REGION Network 14: 关门停止控制
   // 1.脚踢开关又有信号
   // 2.操作门关位有信号
   // 3.操作门关门时间超时
   // 4.门电机保护有信号
   // 5.再次点击开门触摸按钮
   // 6.再次点击关门触摸按钮
   // 7.再次点击机械开门按钮
   // 8.再次点击机械关门按钮
   // 9..操作门有障碍
   RUNG wire#powerrail
      { S7_Templates := "SrcType := Word" } EQ_Contact(in1 := #门状态, in2 := 2)
      wire#w1
      Contact( #脚踢开关状态 )
      wire#w2
      Move(in := 0, out1 => #门状态)
      wire#w3
      R_Coil( #触摸开门按钮状态 )
      R_Coil( #机械开门按钮状态 )
      R_Coil( #机械关门按钮状态 )
      R_Coil( #脚踢开关状态 )
      R_Coil( #触摸关门按钮状态 )
   END_RUNG
   RUNG wire#w1
      Contact( #操作门关位 )
   END_RUNG wire#w2
   RUNG wire#w1
      { S7_Templates := "SrcType := UInt" } GT_Contact(in1 := #关门时间统计, in2 := #操作门最大关闭时间秒)
   END_RUNG wire#w2
   RUNG wire#w1
      Contact( #门电机保护信号 )
   END_RUNG wire#w2
   RUNG wire#w1
      Contact( #机械开门按钮状态 )
   END_RUNG wire#w2
   RUNG wire#w1
      Contact( #机械关门按钮状态 )
   END_RUNG wire#w2
   RUNG wire#w1
      Contact( #触摸关门按钮状态 )
   END_RUNG wire#w2
   RUNG wire#w1
      Contact( #触摸开门按钮状态 )
   END_RUNG wire#w2
   RUNG wire#w1
      I_Contact( #操作门障碍 )
   END_RUNG wire#w2
   RUNG wire#w3
      { S7_Templates := "SrcType := UInt" } GT_Contact(in1 := #关门时间统计, in2 := #操作门最大关闭时间秒)
      I_Contact( #报警开关.%X3 )
      S_Coil( #报警码.%X3 )
   END_RUNG
   RUNG wire#w3
      I_Contact( #操作门障碍 )
      wire#w4
      S_Coil( #关闭门失败后需要开门标志 )
      Move(in := 0, out1 => #门关闭失败重新开门等待时间)
   END_RUNG
   RUNG wire#w4
      I_Contact( #报警开关.%X5 )
      S_Coil( #报警码.%X5 )
   END_RUNG
   RUNG wire#w3
      Contact( #门电机保护信号 )
      I_Contact( #报警开关.%X4 )
      S_Coil( #报警码.%X4 )
   END_RUNG
   // the same network as SCL:
   #_w1 := (#门状态 = 2) AND (#脚踢开关状态 OR #操作门关位 OR (#关门时间统计 > #操作门最大关闭时间秒) OR #门电机保护信号 OR #机械开门按钮状态 OR #机械关门按钮状态 OR #触摸关门按钮状态 OR #触摸开门按钮状态 OR NOT #操作门障碍);
   IF #_w1 THEN
       #门状态 := 0;
       #触摸开门按钮状态 := FALSE;
       #机械开门按钮状态 := FALSE;
       #机械关门按钮状态 := FALSE;
       #脚踢开关状态 := FALSE;
       #触摸关门按钮状态 := FALSE;
   END_IF;
   IF #_w1 AND (#关门时间统计 > #操作门最大关闭时间秒) AND NOT #报警开关.%X3 THEN #报警码.%X3 := TRUE; END_IF;
   #_w2 := #_w1 AND NOT #操作门障碍;
   IF #_w2 THEN
       #关闭门失败后需要开门标志 := TRUE;
       #门关闭失败重新开门等待时间 := 0;
   END_IF;
   IF #_w2 AND NOT #报警开关.%X5 THEN #报警码.%X5 := TRUE; END_IF;
   IF #_w1 AND #门电机保护信号 AND NOT #报警开关.%X4 THEN #报警码.%X4 := TRUE; END_IF;
END_REGION

REGION Network 15: 如果是前门遇到障碍,门停止后,还需要将门打开
   // 关门失败后,门先停止0.8秒 然后再开门
   RUNG wire#powerrail
      { S7_Templates := "SrcType := Word" } EQ_Contact(in1 := #门状态, in2 := 0)
      Contact( #关闭门失败后需要开门标志 )
      wire#w1
      Contact( "Clock_10Hz" )
      P_Trig( #门关闭失败重新开门时间统计沿 )
      { S7_Templates := "DestType := UInt" } Inc( #门关闭失败重新开门等待时间 )
   END_RUNG
   RUNG wire#w1
      { S7_Templates := "SrcType := UInt" } GE_Contact(in1 := #门关闭失败重新开门等待时间, in2 := 8)
      wire#w2
      S_Coil( #触摸开门按钮状态 )
   END_RUNG
   RUNG wire#w2
      R_Coil( #关闭门失败后需要开门标志 )
      Move(in := 0, out1 => #门关闭失败重新开门等待时间)
   END_RUNG
   // the same network as SCL:
   #_w1 := (#门状态 = 0) AND #关闭门失败后需要开门标志;
   #_w2 := #_w1 AND "Clock_10Hz";
   #_w3 := #_w2 AND NOT #门关闭失败重新开门时间统计沿;   // rising edge
   #门关闭失败重新开门时间统计沿 := #_w2;
   IF #_w3 THEN #门关闭失败重新开门等待时间 := #门关闭失败重新开门等待时间 + 1; END_IF;
   IF #_w1 AND (#门关闭失败重新开门等待时间 >= 8) THEN
       #触摸开门按钮状态 := TRUE;
       #关闭门失败后需要开门标志 := FALSE;
       #门关闭失败重新开门等待时间 := 0;
   END_IF;
END_REGION

REGION Network 16: 其他门报警
   // 1.同时检测到操作门关位和开位1秒
   RUNG wire#powerrail
      Contact( #操作门开位 )
      Contact( #操作门关位 )
      wire#w1
      Contact( "Clock_10Hz" )
      P_Trig( #同时检测到门开关位时间统计沿 )
      { S7_Templates := "DestType := UInt" } Inc( #同时检测到门开位和关位信号时间统计 )
   END_RUNG
   RUNG wire#w1
      { S7_Templates := "SrcType := UInt" } GE_Contact(in1 := #同时检测到门开位和关位信号时间统计, in2 := 10)
      Move(in := 10, out1 => #同时检测到门开位和关位信号时间统计)
      I_Contact( #报警开关.%X6 )
      S_Coil( #报警码.%X6 )
   END_RUNG
   RUNG wire#powerrail
      I_Contact( #操作门开位 )
      wire#w2
      Move(in := 0, out1 => #同时检测到门开位和关位信号时间统计)
   END_RUNG
   RUNG wire#powerrail
      I_Contact( #操作门关位 )
   END_RUNG wire#w2
   // the same network as SCL:
   #_w1 := #操作门开位 AND #操作门关位;
   #_w2 := #_w1 AND "Clock_10Hz";
   #_w3 := #_w2 AND NOT #同时检测到门开关位时间统计沿;   // rising edge
   #同时检测到门开关位时间统计沿 := #_w2;
   IF #_w3 THEN #同时检测到门开位和关位信号时间统计 := #同时检测到门开位和关位信号时间统计 + 1; END_IF;
   #_w4 := #_w1 AND (#同时检测到门开位和关位信号时间统计 >= 10);
   IF #_w4 THEN #同时检测到门开位和关位信号时间统计 := 10; END_IF;
   IF #_w4 AND NOT #报警开关.%X6 THEN #报警码.%X6 := TRUE; END_IF;
   IF NOT #操作门开位 OR NOT #操作门关位 THEN #同时检测到门开位和关位信号时间统计 := 0; END_IF;
END_REGION

REGION Network 17: 门运行情况报警码时间统计及清除
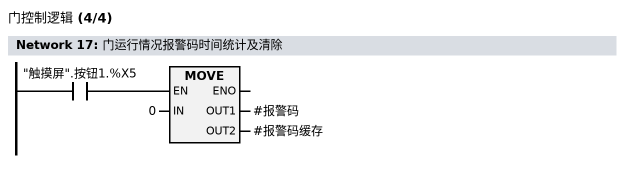
   RUNG wire#powerrail
      Contact( "触摸屏".按钮1.%X5 )
      Move(in := 0, out1 => #报警码, out2 => #报警码缓存)
   END_RUNG
   // the same network as SCL:
   IF "触摸屏".按钮1.%X5 THEN
       #报警码 := 0;
       #报警码缓存 := 0;
   END_IF;
END_REGION
END_FUNCTION_BLOCK

FUNCTION_BLOCK "门功能控制"   // FB15, LAD
{ S7_Optimized_Access := 'TRUE' }
VERSION : 0.1
   VAR_TEMP   // added for the SCL form of the ladder/FBD networks
      _w1 : Bool;
   END_VAR
BEGIN

REGION Network 1
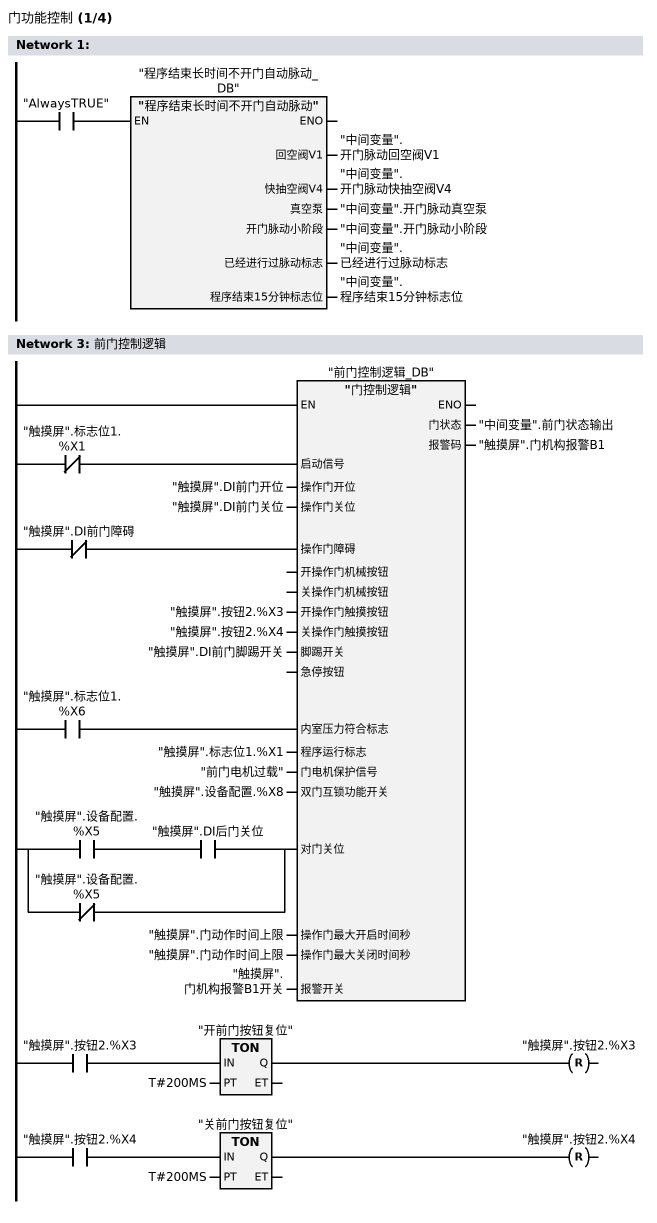
   RUNG wire#powerrail
      Contact( "AlwaysTRUE" )
      "程序结束长时间不开门自动脉动_DB"(回空阀V1 => "中间变量".开门脉动回空阀V1, 快抽空阀V4 => "中间变量".开门脉动快抽空阀V4, 真空泵 => "中间变量".开门脉动真空泵, 开门脉动小阶段 => "中间变量".开门脉动小阶段, 已经进行过脉动标志 => "中间变量".已经进行过脉动标志, 程序结束15分钟标志位 => "中间变量".程序结束15分钟标志位)
   END_RUNG
   // the same network as SCL:
   IF "AlwaysTRUE" THEN
       "程序结束长时间不开门自动脉动_DB"(回空阀V1 => "中间变量".开门脉动回空阀V1,   // "程序结束长时间不开门自动脉动"
                           快抽空阀V4 => "中间变量".开门脉动快抽空阀V4,
                           真空泵 => "中间变量".开门脉动真空泵,
                           开门脉动小阶段 => "中间变量".开门脉动小阶段,
                           已经进行过脉动标志 => "中间变量".已经进行过脉动标志,
                           程序结束15分钟标志位 => "中间变量".程序结束15分钟标志位);
   END_IF;
END_REGION

REGION Network 3: 前门控制逻辑
   "前门控制逻辑_DB"(启动信号 := NOT "触摸屏".标志位1.%X1,   // "门控制逻辑"
               操作门开位 := "触摸屏".DI前门开位,
               操作门关位 := "触摸屏".DI前门关位,
               操作门障碍 := NOT "触摸屏".DI前门障碍,
               开操作门触摸按钮 := "触摸屏".按钮2.%X3,
               关操作门触摸按钮 := "触摸屏".按钮2.%X4,
               脚踢开关 := "触摸屏".DI前门脚踢开关,
               内室压力符合标志 := "触摸屏".标志位1.%X6,
               程序运行标志 := "触摸屏".标志位1.%X1,
               门电机保护信号 := "前门电机过载",
               双门互锁功能开关 := "触摸屏".设备配置.%X8,
               对门关位 := ("触摸屏".设备配置.%X5 AND "触摸屏".DI后门关位) OR NOT "触摸屏".设备配置.%X5,
               操作门最大开启时间秒 := "触摸屏".门动作时间上限,
               操作门最大关闭时间秒 := "触摸屏".门动作时间上限,
               报警开关 := "触摸屏".门机构报警B1开关,
               门状态 => "中间变量".前门状态输出,
               报警码 => "触摸屏".门机构报警B1);
   "开前门按钮复位".TON(IN := "触摸屏".按钮2.%X3, PT := T#200MS);
   IF "开前门按钮复位".Q THEN "触摸屏".按钮2.%X3 := FALSE; END_IF;
   "关前门按钮复位".TON(IN := "触摸屏".按钮2.%X4, PT := T#200MS);
   IF "关前门按钮复位".Q THEN "触摸屏".按钮2.%X4 := FALSE; END_IF;
END_REGION

REGION Network 5: 后门控制逻辑
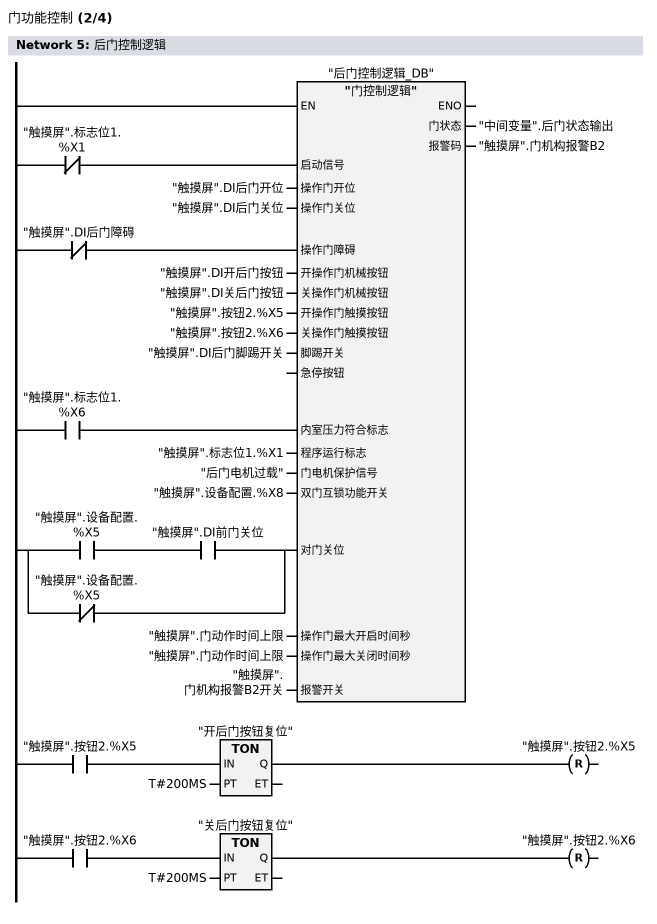
   "后门控制逻辑_DB"(启动信号 := NOT "触摸屏".标志位1.%X1,   // "门控制逻辑"
               操作门开位 := "触摸屏".DI后门开位,
               操作门关位 := "触摸屏".DI后门关位,
               操作门障碍 := NOT "触摸屏".DI后门障碍,
               开操作门机械按钮 := "触摸屏".DI开后门按钮,
               关操作门机械按钮 := "触摸屏".DI关后门按钮,
               开操作门触摸按钮 := "触摸屏".按钮2.%X5,
               关操作门触摸按钮 := "触摸屏".按钮2.%X6,
               脚踢开关 := "触摸屏".DI后门脚踢开关,
               内室压力符合标志 := "触摸屏".标志位1.%X6,
               程序运行标志 := "触摸屏".标志位1.%X1,
               门电机保护信号 := "后门电机过载",
               双门互锁功能开关 := "触摸屏".设备配置.%X8,
               对门关位 := ("触摸屏".设备配置.%X5 AND "触摸屏".DI前门关位) OR NOT "触摸屏".设备配置.%X5,
               操作门最大开启时间秒 := "触摸屏".门动作时间上限,
               操作门最大关闭时间秒 := "触摸屏".门动作时间上限,
               报警开关 := "触摸屏".门机构报警B2开关,
               门状态 => "中间变量".后门状态输出,
               报警码 => "触摸屏".门机构报警B2);
   "开后门按钮复位".TON(IN := "触摸屏".按钮2.%X5, PT := T#200MS);
   IF "开后门按钮复位".Q THEN "触摸屏".按钮2.%X5 := FALSE; END_IF;
   "关后门按钮复位".TON(IN := "触摸屏".按钮2.%X6, PT := T#200MS);
   IF "关后门按钮复位".Q THEN "触摸屏".按钮2.%X6 := FALSE; END_IF;
END_REGION

REGION Network 6: 装载门状态
   // 0故障状态，1前门打开状态后门关闭,2后门打开状态前门关闭，3双门关闭状态，4开前门正在动作，5关前门正在动态，
   // 6开后门正在动作，7关后门正在动作，8门锁紧状态，9两门都开
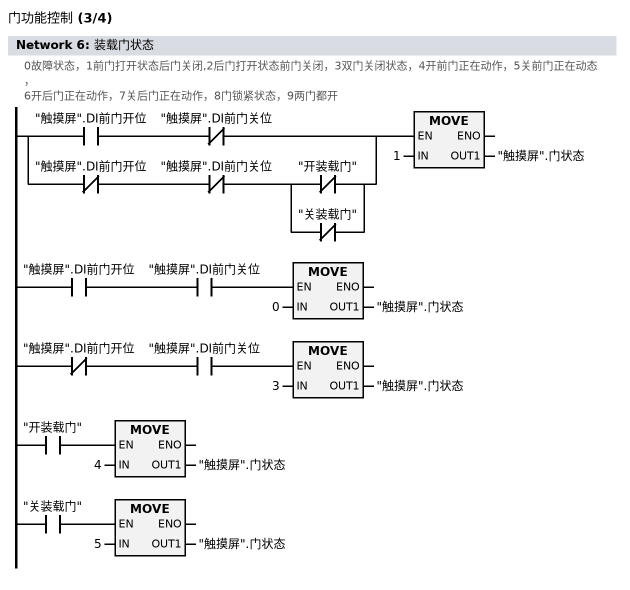
   RUNG wire#powerrail
      Contact( "触摸屏".DI前门开位 )
      I_Contact( "触摸屏".DI前门关位 )
      wire#w1
      Move(in := 1, out1 => "触摸屏".门状态)
   END_RUNG
   RUNG wire#powerrail
      I_Contact( "触摸屏".DI前门开位 )
      I_Contact( "触摸屏".DI前门关位 )
      wire#w2
      I_Contact( "开装载门" )
   END_RUNG wire#w1
   RUNG wire#w2
      I_Contact( "关装载门" )
   END_RUNG wire#w1
   RUNG wire#powerrail
      Contact( "触摸屏".DI前门开位 )
      Contact( "触摸屏".DI前门关位 )
      Move(in := 0, out1 => "触摸屏".门状态)
   END_RUNG
   RUNG wire#powerrail
      I_Contact( "触摸屏".DI前门开位 )
      Contact( "触摸屏".DI前门关位 )
      Move(in := 3, out1 => "触摸屏".门状态)
   END_RUNG
   RUNG wire#powerrail
      Contact( "开装载门" )
      Move(in := 4, out1 => "触摸屏".门状态)
   END_RUNG
   RUNG wire#powerrail
      Contact( "关装载门" )
      Move(in := 5, out1 => "触摸屏".门状态)
   END_RUNG
   // the same network as SCL:
   IF ("触摸屏".DI前门开位 AND NOT "触摸屏".DI前门关位) OR (NOT "触摸屏".DI前门开位 AND NOT "触摸屏".DI前门关位 AND (NOT "开装载门" OR NOT "关装载门")) THEN
       "触摸屏".门状态 := 1;
   END_IF;
   IF "触摸屏".DI前门开位 AND "触摸屏".DI前门关位 THEN "触摸屏".门状态 := 0; END_IF;
   IF NOT "触摸屏".DI前门开位 AND "触摸屏".DI前门关位 THEN "触摸屏".门状态 := 3; END_IF;
   IF "开装载门" THEN "触摸屏".门状态 := 4; END_IF;
   IF "关装载门" THEN "触摸屏".门状态 := 5; END_IF;
END_REGION

REGION Network 7: 卸载门状态
   // 0故障状态，1前门打开状态后门关闭,2后门打开状态前门关闭，3双门关闭状态，4开前门正在动作，5关前门正在动态，
   // 6开后门正在动作，7关后门正在动作，8门锁紧状态，9两门都开
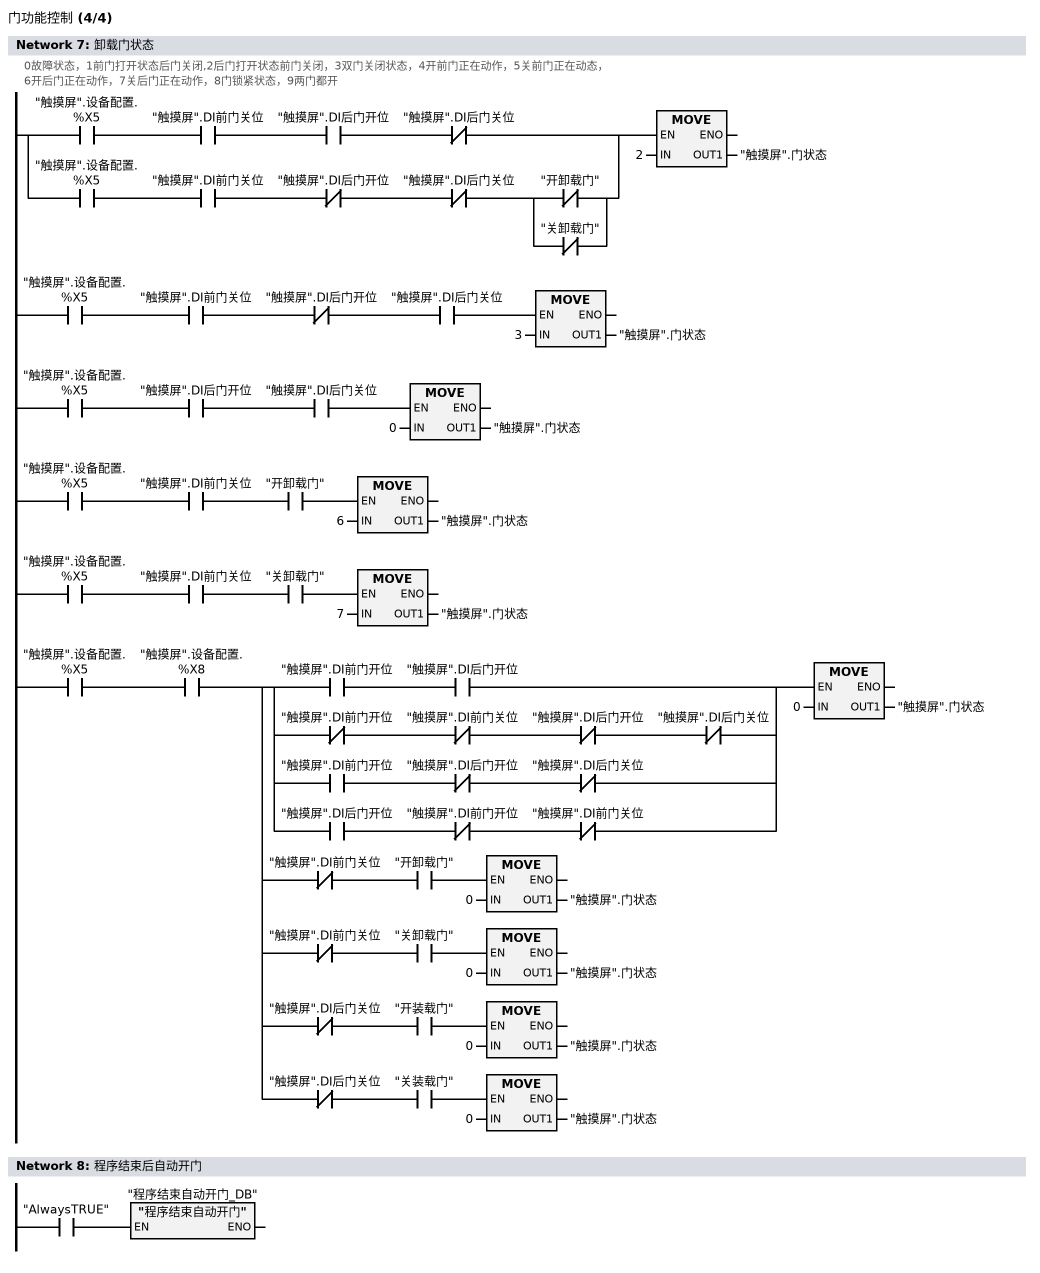
   RUNG wire#powerrail
      Contact( "触摸屏".设备配置.%X5 )
      Contact( "触摸屏".DI前门关位 )
      Contact( "触摸屏".DI后门开位 )
      I_Contact( "触摸屏".DI后门关位 )
      wire#w1
      Move(in := 2, out1 => "触摸屏".门状态)
   END_RUNG
   RUNG wire#powerrail
      Contact( "触摸屏".设备配置.%X5 )
      Contact( "触摸屏".DI前门关位 )
      I_Contact( "触摸屏".DI后门开位 )
      I_Contact( "触摸屏".DI后门关位 )
      wire#w2
      I_Contact( "开卸载门" )
   END_RUNG wire#w1
   RUNG wire#w2
      I_Contact( "关卸载门" )
   END_RUNG wire#w1
   RUNG wire#powerrail
      Contact( "触摸屏".设备配置.%X5 )
      Contact( "触摸屏".DI前门关位 )
      I_Contact( "触摸屏".DI后门开位 )
      Contact( "触摸屏".DI后门关位 )
      Move(in := 3, out1 => "触摸屏".门状态)
   END_RUNG
   RUNG wire#powerrail
      Contact( "触摸屏".设备配置.%X5 )
      Contact( "触摸屏".DI后门开位 )
      Contact( "触摸屏".DI后门关位 )
      Move(in := 0, out1 => "触摸屏".门状态)
   END_RUNG
   RUNG wire#powerrail
      Contact( "触摸屏".设备配置.%X5 )
      Contact( "触摸屏".DI前门关位 )
      Contact( "开卸载门" )
      Move(in := 6, out1 => "触摸屏".门状态)
   END_RUNG
   RUNG wire#powerrail
      Contact( "触摸屏".设备配置.%X5 )
      Contact( "触摸屏".DI前门关位 )
      Contact( "关卸载门" )
      Move(in := 7, out1 => "触摸屏".门状态)
   END_RUNG
   RUNG wire#powerrail
      Contact( "触摸屏".设备配置.%X5 )
      Contact( "触摸屏".设备配置.%X8 )
      wire#w3
      Contact( "触摸屏".DI前门开位 )
      Contact( "触摸屏".DI后门开位 )
      wire#w4
      Move(in := 0, out1 => "触摸屏".门状态)
   END_RUNG
   RUNG wire#w3
      I_Contact( "触摸屏".DI前门开位 )
      I_Contact( "触摸屏".DI前门关位 )
      I_Contact( "触摸屏".DI后门开位 )
      I_Contact( "触摸屏".DI后门关位 )
   END_RUNG wire#w4
   RUNG wire#w3
      Contact( "触摸屏".DI前门开位 )
      I_Contact( "触摸屏".DI后门开位 )
      I_Contact( "触摸屏".DI后门关位 )
   END_RUNG wire#w4
   RUNG wire#w3
      Contact( "触摸屏".DI后门开位 )
      I_Contact( "触摸屏".DI前门开位 )
      I_Contact( "触摸屏".DI前门关位 )
   END_RUNG wire#w4
   RUNG wire#w3
      I_Contact( "触摸屏".DI前门关位 )
      Contact( "开卸载门" )
      Move(in := 0, out1 => "触摸屏".门状态)
   END_RUNG
   RUNG wire#w3
      I_Contact( "触摸屏".DI前门关位 )
      Contact( "关卸载门" )
      Move(in := 0, out1 => "触摸屏".门状态)
   END_RUNG
   RUNG wire#w3
      I_Contact( "触摸屏".DI后门关位 )
      Contact( "开装载门" )
      Move(in := 0, out1 => "触摸屏".门状态)
   END_RUNG
   RUNG wire#w3
      I_Contact( "触摸屏".DI后门关位 )
      Contact( "关装载门" )
      Move(in := 0, out1 => "触摸屏".门状态)
   END_RUNG
   // the same network as SCL:
   IF ("触摸屏".设备配置.%X5 AND "触摸屏".DI前门关位 AND "触摸屏".DI后门开位 AND NOT "触摸屏".DI后门关位) OR ("触摸屏".设备配置.%X5 AND "触摸屏".DI前门关位 AND NOT "触摸屏".DI后门开位 AND NOT "触摸屏".DI后门关位 AND (NOT "开卸载门" OR NOT "关卸载门")) THEN
       "触摸屏".门状态 := 2;
   END_IF;
   IF "触摸屏".设备配置.%X5 AND "触摸屏".DI前门关位 AND NOT "触摸屏".DI后门开位 AND "触摸屏".DI后门关位 THEN "触摸屏".门状态 := 3; END_IF;
   IF "触摸屏".设备配置.%X5 AND "触摸屏".DI后门开位 AND "触摸屏".DI后门关位 THEN "触摸屏".门状态 := 0; END_IF;
   IF "触摸屏".设备配置.%X5 AND "触摸屏".DI前门关位 AND "开卸载门" THEN "触摸屏".门状态 := 6; END_IF;
   IF "触摸屏".设备配置.%X5 AND "触摸屏".DI前门关位 AND "关卸载门" THEN "触摸屏".门状态 := 7; END_IF;
   #_w1 := "触摸屏".设备配置.%X5 AND "触摸屏".设备配置.%X8;
   IF #_w1 AND (("触摸屏".DI前门开位 AND "触摸屏".DI后门开位) OR (NOT "触摸屏".DI前门开位 AND NOT "触摸屏".DI前门关位 AND NOT "触摸屏".DI后门开位 AND NOT "触摸屏".DI后门关位) OR ("触摸屏".DI前门开位 AND NOT "触摸屏".DI后门开位 AND NOT "触摸屏".DI后门关位) OR ("触摸屏".DI后门开位 AND NOT "触摸屏".DI前门开位 AND NOT "触摸屏".DI前门关位)) THEN
       "触摸屏".门状态 := 0;
   END_IF;
   IF #_w1 AND NOT "触摸屏".DI前门关位 AND "开卸载门" THEN "触摸屏".门状态 := 0; END_IF;
   IF #_w1 AND NOT "触摸屏".DI前门关位 AND "关卸载门" THEN "触摸屏".门状态 := 0; END_IF;
   IF #_w1 AND NOT "触摸屏".DI后门关位 AND "开装载门" THEN "触摸屏".门状态 := 0; END_IF;
   IF #_w1 AND NOT "触摸屏".DI后门关位 AND "关装载门" THEN "触摸屏".门状态 := 0; END_IF;
END_REGION

REGION Network 8: 程序结束后自动开门
   RUNG wire#powerrail
      Contact( "AlwaysTRUE" )
      "程序结束自动开门_DB"()
   END_RUNG
   // the same network as SCL:
   IF "AlwaysTRUE" THEN
       "程序结束自动开门_DB"();   // "程序结束自动开门"
   END_IF;
END_REGION
END_FUNCTION_BLOCK

FUNCTION_BLOCK "程序结束自动开门"   // FB25, LAD
{ S7_Optimized_Access := 'TRUE' }
VERSION : 0.1
// 自动开门的小阶段
   VAR
      自动开门小阶段 : Int;
   END_VAR
   VAR_TEMP   // added for the SCL form of the ladder/FBD networks
      _w1 : Bool;
   END_VAR
BEGIN

REGION Network 1: 待机阶段
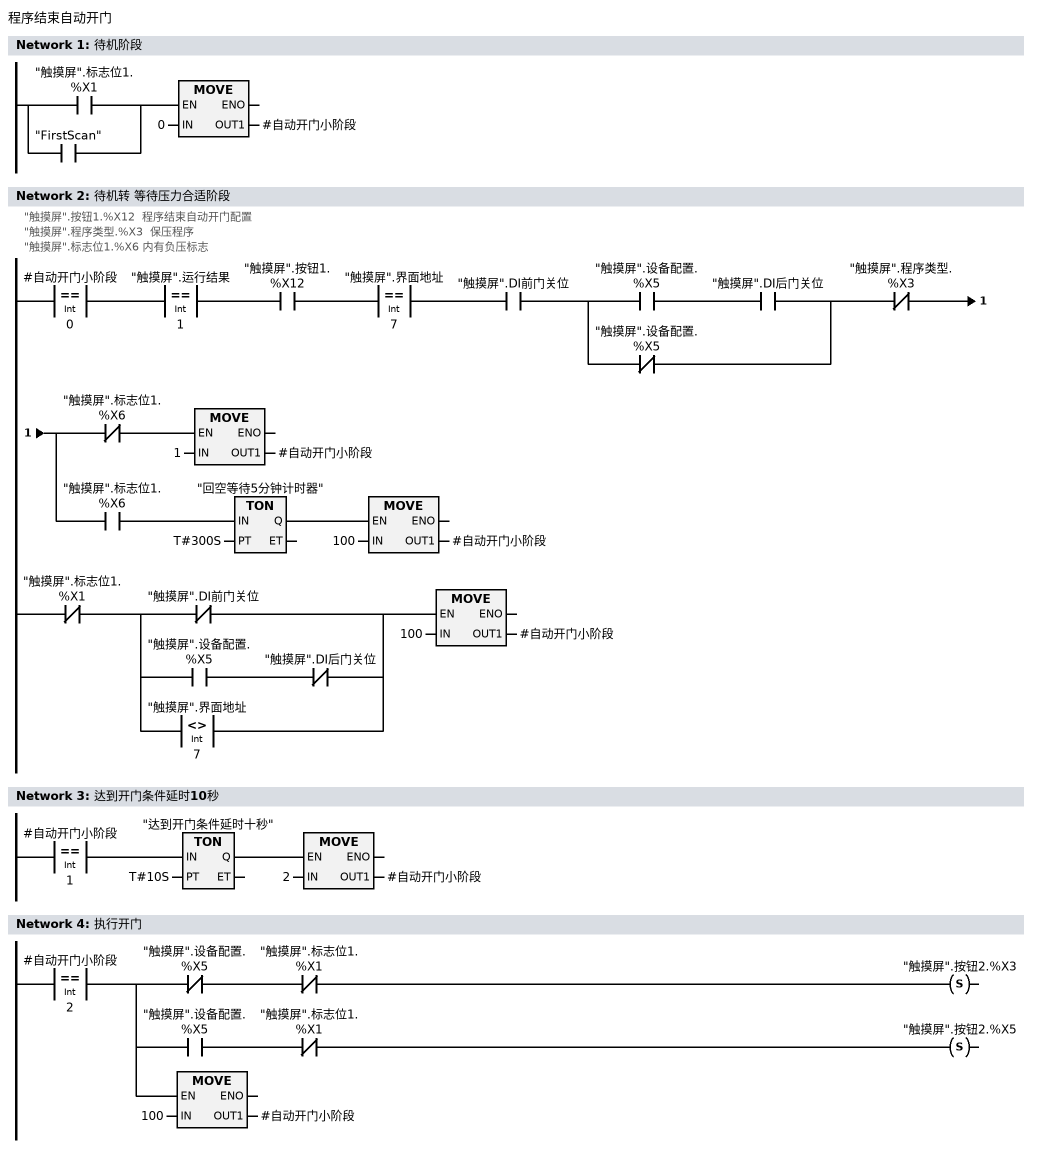
   RUNG wire#powerrail
      Contact( "触摸屏".标志位1.%X1 )
      wire#w1
      { S7_GenerateENO := "TRUE" } Move(in := 0, out1 => #自动开门小阶段)
   END_RUNG
   RUNG wire#powerrail
      Contact( "FirstScan" )
   END_RUNG wire#w1
   // the same network as SCL:
   IF "触摸屏".标志位1.%X1 OR "FirstScan" THEN #自动开门小阶段 := 0; END_IF;
END_REGION

REGION Network 2: 待机转 等待压力合适阶段
   // "触摸屏".按钮1.%X12  程序结束自动开门配置 
   // "触摸屏".程序类型.%X3  保压程序
   // "触摸屏".标志位1.%X6 内有负压标志
   #_w1 := (#自动开门小阶段 = 0) AND ("触摸屏".运行结果 = 1) AND "触摸屏".按钮1.%X12 AND ("触摸屏".界面地址 = 7) AND "触摸屏".DI前门关位 AND (("触摸屏".设备配置.%X5 AND "触摸屏".DI后门关位) OR NOT "触摸屏".设备配置.%X5) AND NOT "触摸屏".程序类型.%X3;
   IF #_w1 AND NOT "触摸屏".标志位1.%X6 THEN #自动开门小阶段 := 1; END_IF;
   "回空等待5分钟计时器".TON(IN := #_w1 AND "触摸屏".标志位1.%X6, PT := T#300S);
   IF "回空等待5分钟计时器".Q THEN #自动开门小阶段 := 100; END_IF;
   IF NOT "触摸屏".标志位1.%X1 AND (NOT "触摸屏".DI前门关位 OR ("触摸屏".设备配置.%X5 AND NOT "触摸屏".DI后门关位) OR ("触摸屏".界面地址 <> 7)) THEN
       #自动开门小阶段 := 100;
   END_IF;
END_REGION

REGION Network 3: 达到开门条件延时10秒
   "达到开门条件延时十秒".TON(IN := #自动开门小阶段 = 1, PT := T#10S);
   IF "达到开门条件延时十秒".Q THEN #自动开门小阶段 := 2; END_IF;
END_REGION

REGION Network 4: 执行开门
   RUNG wire#powerrail
      { S7_Templates := "SrcType := Int" } EQ_Contact(in1 := #自动开门小阶段, in2 := 2)
      wire#w1
      I_Contact( "触摸屏".设备配置.%X5 )
      I_Contact( "触摸屏".标志位1.%X1 )
      S_Coil( "触摸屏".按钮2.%X3 )
   END_RUNG
   RUNG wire#w1
      Contact( "触摸屏".设备配置.%X5 )
      I_Contact( "触摸屏".标志位1.%X1 )
      S_Coil( "触摸屏".按钮2.%X5 )
   END_RUNG
   RUNG wire#w1
      { S7_GenerateENO := "TRUE" } Move(in := 100, out1 => #自动开门小阶段)
   END_RUNG
   // the same network as SCL:
   #_w1 := #自动开门小阶段 = 2;
   IF #_w1 AND NOT "触摸屏".设备配置.%X5 AND NOT "触摸屏".标志位1.%X1 THEN "触摸屏".按钮2.%X3 := TRUE; END_IF;
   IF #_w1 AND "触摸屏".设备配置.%X5 AND NOT "触摸屏".标志位1.%X1 THEN "触摸屏".按钮2.%X5 := TRUE; END_IF;
   IF #_w1 THEN #自动开门小阶段 := 100; END_IF;
END_REGION

REGION Network 5: 结束 100
END_REGION
END_FUNCTION_BLOCK

FUNCTION_BLOCK "程序结束长时间不开门自动脉动"   // FB26, LAD
{ S7_Optimized_Access := 'TRUE' }
VERSION : 0.1
   VAR_OUTPUT
      回空阀V1 : Bool;
      快抽空阀V4 : Bool;
      真空泵 : Bool;
      开门脉动小阶段 : Int;
      已经进行过脉动标志 : Int;
      程序结束15分钟标志位 : Int;
   END_VAR
   VAR RETAIN
      正在进行开门脉动标志 : Int;
      已进行过开门脉动标志 : Int;
      程序结束15分钟标志 : Int;
      结束满足压力 : Int;
      开门触发的位置 : Int;
      程序正常结束标志 : Bool;
   END_VAR
   VAR_TEMP   // added for the SCL form of the ladder/FBD networks
      _w1 : Bool;
   END_VAR
BEGIN

REGION Network 1: 待机阶段
   // 开门脉动小阶段：0未进行 1抽空 2回空 3结束
   // 正在进行开门脉动标志：0未进行 1正在进行
   // 已进行过开门脉动标志：0未进行 1已经进行
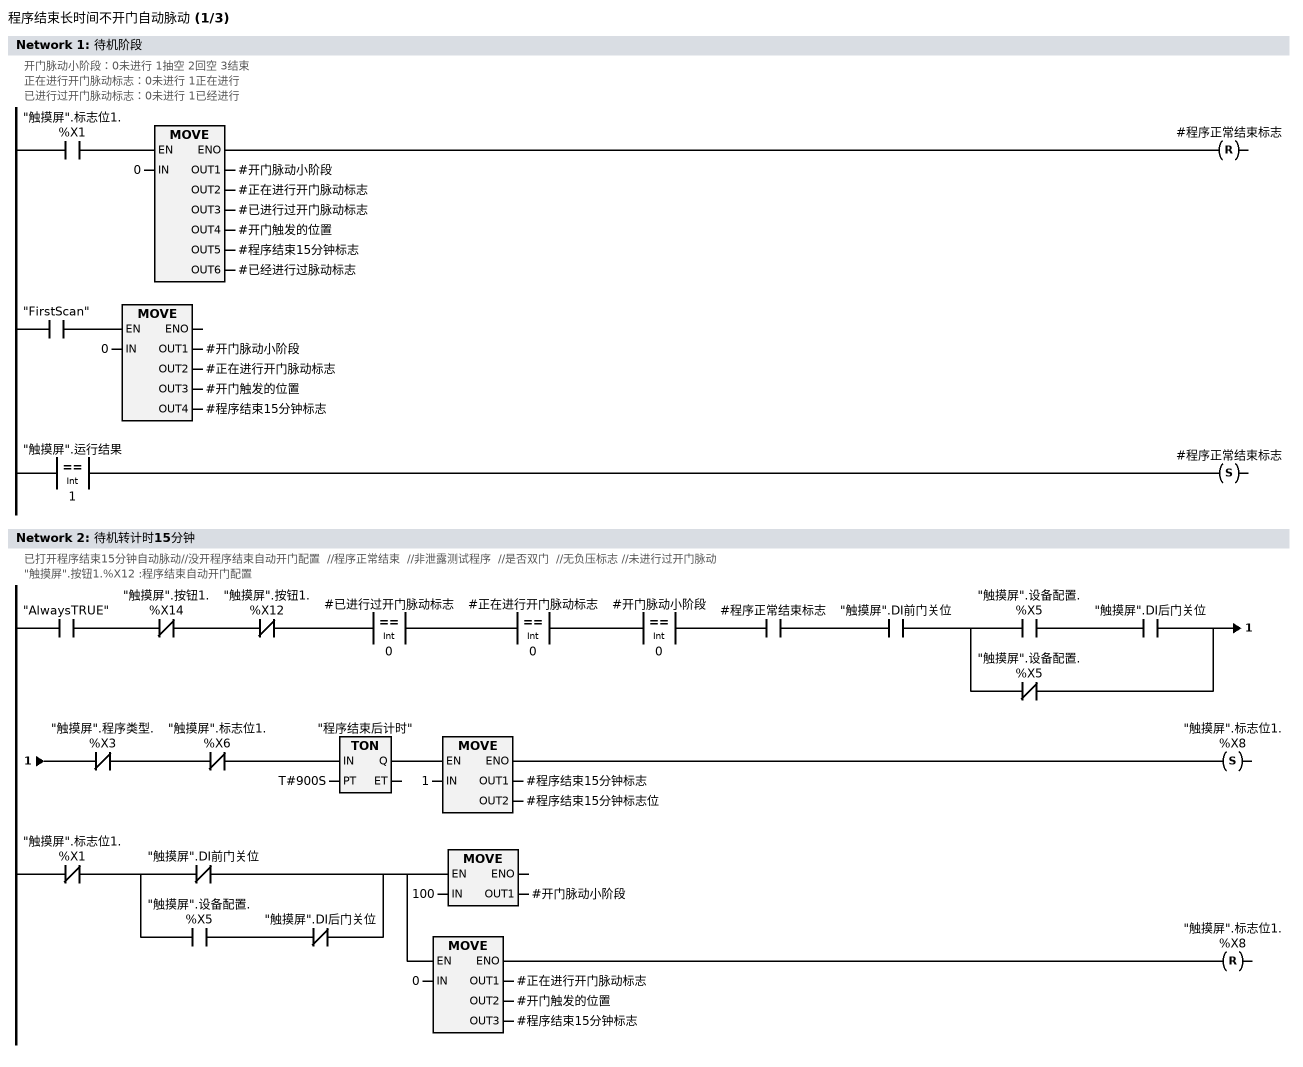
   RUNG wire#powerrail
      Contact( "触摸屏".标志位1.%X1 )
      { S7_GenerateENO := "TRUE" } Move(in := 0, out1 => #开门脉动小阶段, out2 => #正在进行开门脉动标志, out3 => #已进行过开门脉动标志, out4 => #开门触发的位置, out5 => #程序结束15分钟标志, out6 => #已经进行过脉动标志)
      R_Coil( #程序正常结束标志 )
   END_RUNG
   RUNG wire#powerrail
      Contact( "FirstScan" )
      { S7_GenerateENO := "TRUE" } Move(in := 0, out1 => #开门脉动小阶段, out2 => #正在进行开门脉动标志, out3 => #开门触发的位置, out4 => #程序结束15分钟标志)
   END_RUNG
   RUNG wire#powerrail
      { S7_Templates := "SrcType := Int" } EQ_Contact(in1 := "触摸屏".运行结果, in2 := 1)
      S_Coil( #程序正常结束标志 )
   END_RUNG
   // the same network as SCL:
   // ENO of a box is taken as its EN; it also drops when the box reports an error
   IF "触摸屏".标志位1.%X1 THEN
       #开门脉动小阶段 := 0;
       #正在进行开门脉动标志 := 0;
       #已进行过开门脉动标志 := 0;
       #开门触发的位置 := 0;
       #程序结束15分钟标志 := 0;
       #已经进行过脉动标志 := 0;
       #程序正常结束标志 := FALSE;
   END_IF;
   IF "FirstScan" THEN
       #开门脉动小阶段 := 0;
       #正在进行开门脉动标志 := 0;
       #开门触发的位置 := 0;
       #程序结束15分钟标志 := 0;
   END_IF;
   IF "触摸屏".运行结果 = 1 THEN #程序正常结束标志 := TRUE; END_IF;
END_REGION

REGION Network 2: 待机转计时15分钟
   // 已打开程序结束15分钟自动脉动//没开程序结束自动开门配置  //程序正常结束  //非泄露测试程序  //是否双门  //无负压标志 //未进行过开门脉动
   // "触摸屏".按钮1.%X12 :程序结束自动开门配置
   // ENO of a box is taken as its EN; it also drops when the box reports an error
   "程序结束后计时".TON(IN := "AlwaysTRUE" AND NOT "触摸屏".按钮1.%X14 AND NOT "触摸屏".按钮1.%X12 AND (#已进行过开门脉动标志 = 0) AND (#正在进行开门脉动标志 = 0) AND (#开门脉动小阶段 = 0) AND #程序正常结束标志 AND "触摸屏".DI前门关位 AND (("触摸屏".设备配置.%X5 AND "触摸屏".DI后门关位) OR NOT "触摸屏".设备配置.%X5) AND NOT "触摸屏".程序类型.%X3 AND NOT "触摸屏".标志位1.%X6,
                 PT := T#900S);
   IF "程序结束后计时".Q THEN
       #程序结束15分钟标志 := 1;
       #程序结束15分钟标志位 := 1;
       "触摸屏".标志位1.%X8 := TRUE;
   END_IF;
   IF NOT "触摸屏".标志位1.%X1 AND (NOT "触摸屏".DI前门关位 OR ("触摸屏".设备配置.%X5 AND NOT "触摸屏".DI后门关位)) THEN
       #开门脉动小阶段 := 100;
       #正在进行开门脉动标志 := 0;
       #开门触发的位置 := 0;
       #程序结束15分钟标志 := 0;
       "触摸屏".标志位1.%X8 := FALSE;
   END_IF;
END_REGION

REGION Network 3: 保存 开门触发的位置
   // 开门触发的位置:0未触发 1开装载门按钮 2装载门脚踢 3开卸载门物理按钮 4卸载门脚踢 5开卸载门按钮
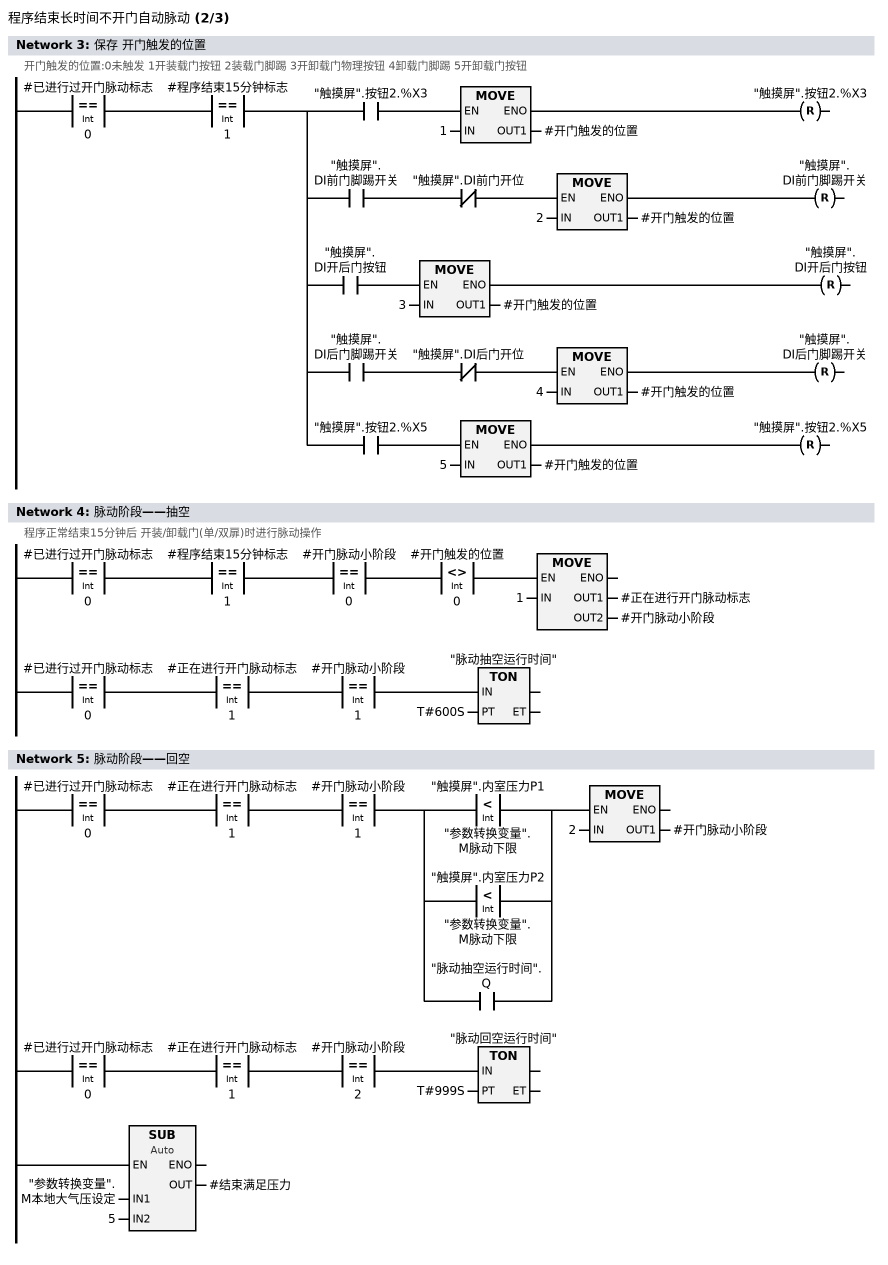
   RUNG wire#powerrail
      { S7_Templates := "SrcType := Int" } EQ_Contact(in1 := #已进行过开门脉动标志, in2 := 0)
      { S7_Templates := "SrcType := Int" } EQ_Contact(in1 := #程序结束15分钟标志, in2 := 1)
      wire#w1
      Contact( "触摸屏".按钮2.%X3 )
      { S7_GenerateENO := "TRUE" } Move(in := 1, out1 => #开门触发的位置)
      R_Coil( "触摸屏".按钮2.%X3 )
   END_RUNG
   RUNG wire#w1
      Contact( "触摸屏".DI前门脚踢开关 )
      I_Contact( "触摸屏".DI前门开位 )
      { S7_GenerateENO := "TRUE" } Move(in := 2, out1 => #开门触发的位置)
      R_Coil( "触摸屏".DI前门脚踢开关 )
   END_RUNG
   RUNG wire#w1
      Contact( "触摸屏".DI开后门按钮 )
      { S7_GenerateENO := "TRUE" } Move(in := 3, out1 => #开门触发的位置)
      R_Coil( "触摸屏".DI开后门按钮 )
   END_RUNG
   RUNG wire#w1
      Contact( "触摸屏".DI后门脚踢开关 )
      I_Contact( "触摸屏".DI后门开位 )
      { S7_GenerateENO := "TRUE" } Move(in := 4, out1 => #开门触发的位置)
      R_Coil( "触摸屏".DI后门脚踢开关 )
   END_RUNG
   RUNG wire#w1
      Contact( "触摸屏".按钮2.%X5 )
      { S7_GenerateENO := "TRUE" } Move(in := 5, out1 => #开门触发的位置)
      R_Coil( "触摸屏".按钮2.%X5 )
   END_RUNG
   // the same network as SCL:
   // ENO of a box is taken as its EN; it also drops when the box reports an error
   #_w1 := (#已进行过开门脉动标志 = 0) AND (#程序结束15分钟标志 = 1);
   IF #_w1 AND "触摸屏".按钮2.%X3 THEN
       #开门触发的位置 := 1;
       "触摸屏".按钮2.%X3 := FALSE;
   END_IF;
   IF #_w1 AND "触摸屏".DI前门脚踢开关 AND NOT "触摸屏".DI前门开位 THEN
       #开门触发的位置 := 2;
       "触摸屏".DI前门脚踢开关 := FALSE;
   END_IF;
   IF #_w1 AND "触摸屏".DI开后门按钮 THEN
       #开门触发的位置 := 3;
       "触摸屏".DI开后门按钮 := FALSE;
   END_IF;
   IF #_w1 AND "触摸屏".DI后门脚踢开关 AND NOT "触摸屏".DI后门开位 THEN
       #开门触发的位置 := 4;
       "触摸屏".DI后门脚踢开关 := FALSE;
   END_IF;
   IF #_w1 AND "触摸屏".按钮2.%X5 THEN
       #开门触发的位置 := 5;
       "触摸屏".按钮2.%X5 := FALSE;
   END_IF;
END_REGION

REGION Network 4: 脉动阶段——抽空
   // 程序正常结束15分钟后 开装/卸载门(单/双扉)时进行脉动操作
   IF (#已进行过开门脉动标志 = 0) AND (#程序结束15分钟标志 = 1) AND (#开门脉动小阶段 = 0) AND (#开门触发的位置 <> 0) THEN
       #正在进行开门脉动标志 := 1;
       #开门脉动小阶段 := 1;
   END_IF;
   "脉动抽空运行时间".TON(IN := (#已进行过开门脉动标志 = 0) AND (#正在进行开门脉动标志 = 1) AND (#开门脉动小阶段 = 1), PT := T#600S);
END_REGION

REGION Network 5: 脉动阶段——回空
   IF (#已进行过开门脉动标志 = 0) AND (#正在进行开门脉动标志 = 1) AND (#开门脉动小阶段 = 1) AND (("触摸屏".内室压力P1 < "参数转换变量".M脉动下限) OR ("触摸屏".内室压力P2 < "参数转换变量".M脉动下限) OR "脉动抽空运行时间".Q) THEN
       #开门脉动小阶段 := 2;
   END_IF;
   "脉动回空运行时间".TON(IN := (#已进行过开门脉动标志 = 0) AND (#正在进行开门脉动标志 = 1) AND (#开门脉动小阶段 = 2), PT := T#999S);
   #结束满足压力 := "参数转换变量".M本地大气压设定 - 5;
END_REGION

REGION Network 6: 脉动阶段——结束
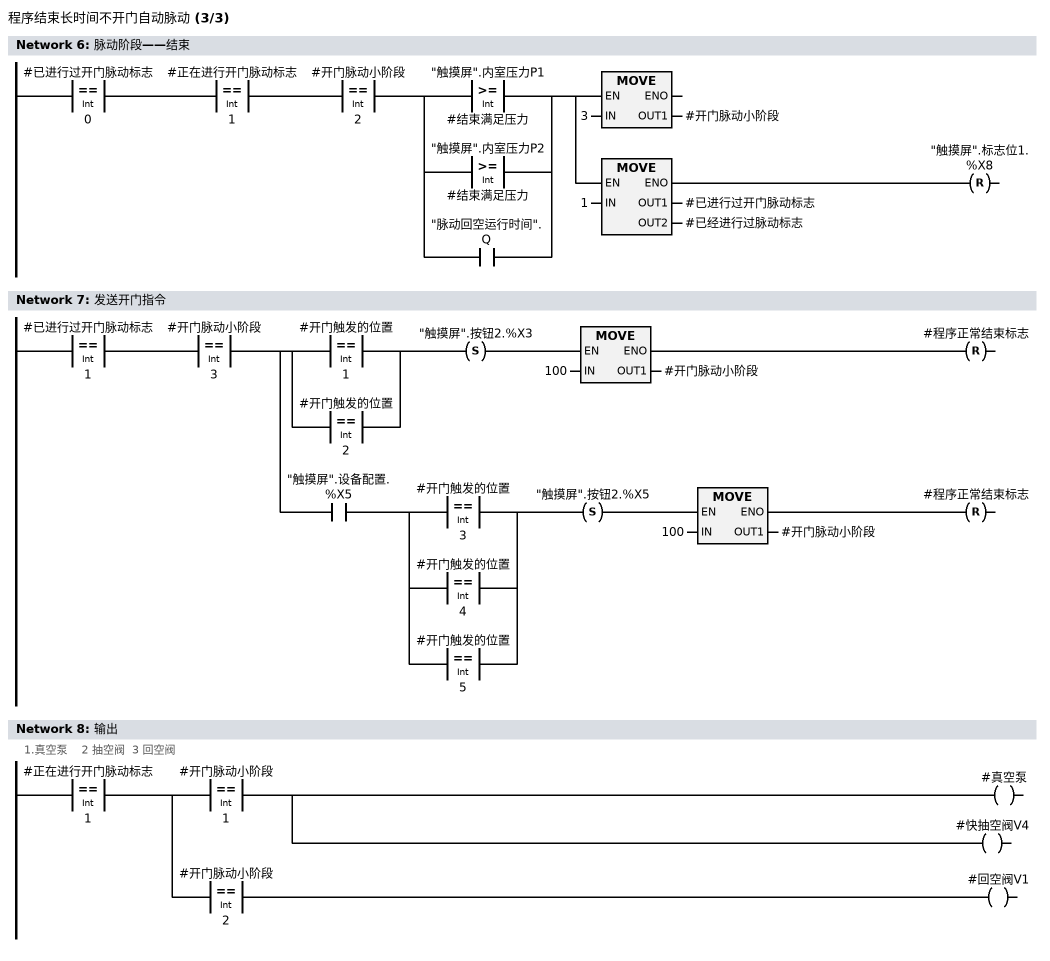
   RUNG wire#powerrail
      { S7_Templates := "SrcType := Int" } EQ_Contact(in1 := #已进行过开门脉动标志, in2 := 0)
      { S7_Templates := "SrcType := Int" } EQ_Contact(in1 := #正在进行开门脉动标志, in2 := 1)
      { S7_Templates := "SrcType := Int" } EQ_Contact(in1 := #开门脉动小阶段, in2 := 2)
      wire#w1
      { S7_Templates := "SrcType := Int" } GE_Contact(in1 := "触摸屏".内室压力P1, in2 := #结束满足压力)
      wire#w2
      { S7_GenerateENO := "TRUE" } Move(in := 3, out1 => #开门脉动小阶段)
   END_RUNG
   RUNG wire#w1
      { S7_Templates := "SrcType := Int" } GE_Contact(in1 := "触摸屏".内室压力P2, in2 := #结束满足压力)
   END_RUNG wire#w2
   RUNG wire#w1
      Contact( "脉动回空运行时间".Q )
   END_RUNG wire#w2
   RUNG wire#w2
      { S7_GenerateENO := "TRUE" } Move(in := 1, out1 => #已进行过开门脉动标志, out2 => #已经进行过脉动标志)
      R_Coil( "触摸屏".标志位1.%X8 )
   END_RUNG
   // the same network as SCL:
   // ENO of a box is taken as its EN; it also drops when the box reports an error
   #_w1 := (#已进行过开门脉动标志 = 0) AND (#正在进行开门脉动标志 = 1) AND (#开门脉动小阶段 = 2) AND (("触摸屏".内室压力P1 >= #结束满足压力) OR ("触摸屏".内室压力P2 >= #结束满足压力) OR "脉动回空运行时间".Q);
   IF #_w1 THEN
       #开门脉动小阶段 := 3;
       #已进行过开门脉动标志 := 1;
       #已经进行过脉动标志 := 1;
       "触摸屏".标志位1.%X8 := FALSE;
   END_IF;
END_REGION

REGION Network 7: 发送开门指令
   RUNG wire#powerrail
      { S7_Templates := "SrcType := Int" } EQ_Contact(in1 := #已进行过开门脉动标志, in2 := 1)
      { S7_Templates := "SrcType := Int" } EQ_Contact(in1 := #开门脉动小阶段, in2 := 3)
      wire#w1
      { S7_Templates := "SrcType := Int" } EQ_Contact(in1 := #开门触发的位置, in2 := 1)
      wire#w2
      S_Coil( "触摸屏".按钮2.%X3 )
      { S7_GenerateENO := "TRUE" } Move(in := 100, out1 => #开门脉动小阶段)
      R_Coil( #程序正常结束标志 )
   END_RUNG
   RUNG wire#w1
      { S7_Templates := "SrcType := Int" } EQ_Contact(in1 := #开门触发的位置, in2 := 2)
   END_RUNG wire#w2
   RUNG wire#w1
      Contact( "触摸屏".设备配置.%X5 )
      wire#w3
      { S7_Templates := "SrcType := Int" } EQ_Contact(in1 := #开门触发的位置, in2 := 3)
      wire#w4
      S_Coil( "触摸屏".按钮2.%X5 )
      { S7_GenerateENO := "TRUE" } Move(in := 100, out1 => #开门脉动小阶段)
      R_Coil( #程序正常结束标志 )
   END_RUNG
   RUNG wire#w3
      { S7_Templates := "SrcType := Int" } EQ_Contact(in1 := #开门触发的位置, in2 := 4)
   END_RUNG wire#w4
   RUNG wire#w3
      { S7_Templates := "SrcType := Int" } EQ_Contact(in1 := #开门触发的位置, in2 := 5)
   END_RUNG wire#w4
   // the same network as SCL:
   // ENO of a box is taken as its EN; it also drops when the box reports an error
   #_w1 := (#已进行过开门脉动标志 = 1) AND (#开门脉动小阶段 = 3);
   IF #_w1 AND ((#开门触发的位置 = 1) OR (#开门触发的位置 = 2)) THEN
       "触摸屏".按钮2.%X3 := TRUE;
       #开门脉动小阶段 := 100;
       #程序正常结束标志 := FALSE;
   END_IF;
   IF #_w1 AND "触摸屏".设备配置.%X5 AND ((#开门触发的位置 = 3) OR (#开门触发的位置 = 4) OR (#开门触发的位置 = 5)) THEN
       "触摸屏".按钮2.%X5 := TRUE;
       #开门脉动小阶段 := 100;
       #程序正常结束标志 := FALSE;
   END_IF;
END_REGION

REGION Network 8: 输出
   // 1.真空泵    2 抽空阀  3 回空阀
   RUNG wire#powerrail
      { S7_Templates := "SrcType := Int" } EQ_Contact(in1 := #正在进行开门脉动标志, in2 := 1)
      wire#w1
      { S7_Templates := "SrcType := Int" } EQ_Contact(in1 := #开门脉动小阶段, in2 := 1)
      wire#w2
      Coil( #真空泵 )
   END_RUNG
   RUNG wire#w2
      Coil( #快抽空阀V4 )
   END_RUNG
   RUNG wire#w1
      { S7_Templates := "SrcType := Int" } EQ_Contact(in1 := #开门脉动小阶段, in2 := 2)
      Coil( #回空阀V1 )
   END_RUNG
   // the same network as SCL:
   #_w1 := #正在进行开门脉动标志 = 1;
   #真空泵 := #_w1 AND (#开门脉动小阶段 = 1);
   #快抽空阀V4 := #真空泵;
   #回空阀V1 := #_w1 AND (#开门脉动小阶段 = 2);
END_REGION
END_FUNCTION_BLOCK

// folder: 14加热功能控制

FUNCTION_BLOCK "加热功能控制"   // FB18, LAD
{ S7_Optimized_Access := 'TRUE' }
VERSION : 0.1
   VAR
      中间变量 : Int;
      催化加热温度上限 : Int;
      催化箱加热标志 : Bool;
      汽化器加热下限 : Int;
      汽化器加热标志 : Bool;
      汽化器加热上限 : Int;
      湿化汽化器加热下限 : Int;
      湿化汽化器加热上限 : Int;
      开始加热下限 : Int;
      前部加热下限 : Int;
      前部加热上限 : Int;
      前部加热标志 : Bool;
      后部加热下限 : Int;
      后部加热上限 : Int;
      后部加热标志 : Bool;
      后门加热下限 : Int;
      后门加热上限 : Int;
      后门加热标志 : Bool;
      前门加热下限 : Int;
      前门加热上限 : Int;
      前门加热标志 : Bool;
      前部停止加热上限 : Int;
      后部停止加热上限 : Int;
      前门停止加热上限 : Int;
      后门停止加热上限 : Int;
      前部启动加热上限 : Int;
      后部启动加热上限 : Int;
      前门启动加热上限 : Int;
      后门启动加热上限 : Int;
      前部启动加热下限 : Int;
      后部启动加热下限 : Int;
      前门启动加热下限 : Int;
      后门启动加热下限 : Int;
      腔体前部加热计时秒 : Int;
      汽化器加热计时秒 : Int;
      腔体后部加热计时秒 : Int;
      前门加热计时秒 : Int;
      后门加热计时秒 : Int;
      催化箱加热计时秒 : Int;
      沿1 : Bool;
      沿2 : Bool;
      沿3 : Bool;
      沿4 : Bool;
      沿5 : Bool;
   END_VAR
   VAR_TEMP   // added for the SCL form of the ladder/FBD networks
      _w1 : Bool;
      _w2 : Bool;
      _w3 : Bool;
   END_VAR
BEGIN

REGION Network 1: 催化箱加热控制
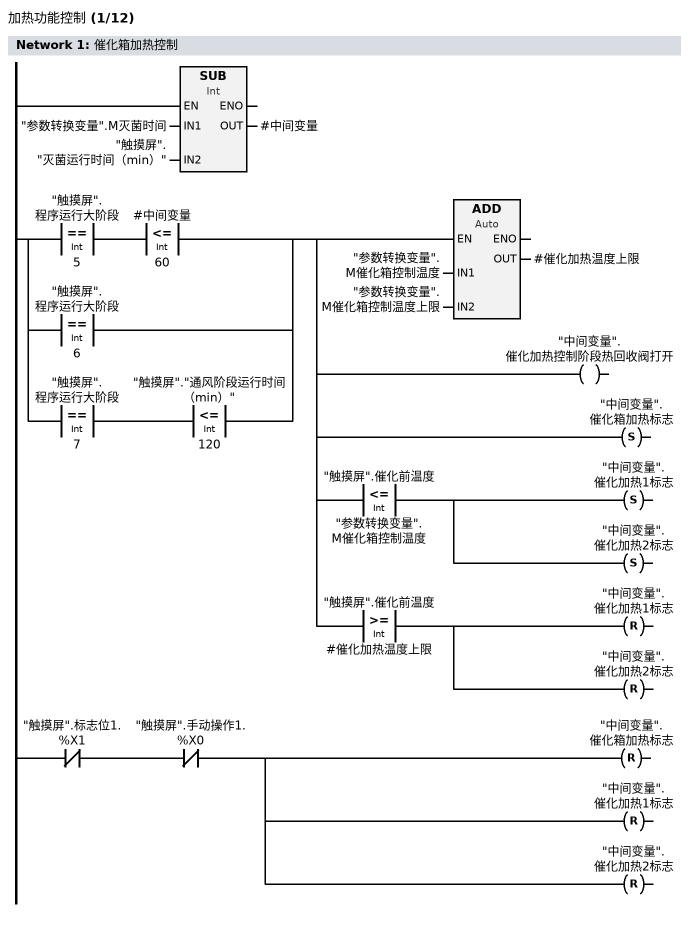
   RUNG wire#powerrail
      { S7_Templates := "SrcType := Int" } Sub(in1 := "参数转换变量".M灭菌时间, in2 := "触摸屏"."灭菌运行时间（min）", out => #中间变量)
   END_RUNG
   RUNG wire#powerrail
      { S7_Templates := "SrcType := Int" } EQ_Contact(in1 := "触摸屏".程序运行大阶段, in2 := 5)
      { S7_Templates := "SrcType := Int" } LE_Contact(in1 := #中间变量, in2 := 60)
      wire#w1
      Add(in1 := "参数转换变量".M催化箱控制温度, in2 := "参数转换变量".M催化箱控制温度上限, out => #催化加热温度上限)
   END_RUNG
   RUNG wire#powerrail
      { S7_Templates := "SrcType := Int" } EQ_Contact(in1 := "触摸屏".程序运行大阶段, in2 := 6)
   END_RUNG wire#w1
   RUNG wire#powerrail
      { S7_Templates := "SrcType := Int" } EQ_Contact(in1 := "触摸屏".程序运行大阶段, in2 := 7)
      { S7_Templates := "SrcType := Int" } LE_Contact(in1 := "触摸屏"."通风阶段运行时间（min）", in2 := 120)
   END_RUNG wire#w1
   RUNG wire#w1
      Coil( "中间变量".催化加热控制阶段热回收阀打开 )
   END_RUNG
   RUNG wire#w1
      S_Coil( "中间变量".催化箱加热标志 )
   END_RUNG
   RUNG wire#w1
      { S7_Templates := "SrcType := Int" } LE_Contact(in1 := "触摸屏".催化前温度, in2 := "参数转换变量".M催化箱控制温度)
      wire#w2
      S_Coil( "中间变量".催化加热1标志 )
   END_RUNG
   RUNG wire#w2
      S_Coil( "中间变量".催化加热2标志 )
   END_RUNG
   RUNG wire#w1
      { S7_Templates := "SrcType := Int" } GE_Contact(in1 := "触摸屏".催化前温度, in2 := #催化加热温度上限)
      wire#w3
      R_Coil( "中间变量".催化加热1标志 )
   END_RUNG
   RUNG wire#w3
      R_Coil( "中间变量".催化加热2标志 )
   END_RUNG
   RUNG wire#powerrail
      I_Contact( "触摸屏".标志位1.%X1 )
      I_Contact( "触摸屏".手动操作1.%X0 )
      wire#w4
      R_Coil( "中间变量".催化箱加热标志 )
   END_RUNG
   RUNG wire#w4
      R_Coil( "中间变量".催化加热1标志 )
   END_RUNG
   RUNG wire#w4
      R_Coil( "中间变量".催化加热2标志 )
   END_RUNG
   // the same network as SCL:
   #中间变量 := "参数转换变量".M灭菌时间 - "触摸屏"."灭菌运行时间（min）";
   #_w1 := (("触摸屏".程序运行大阶段 = 5) AND (#中间变量 <= 60)) OR ("触摸屏".程序运行大阶段 = 6) OR (("触摸屏".程序运行大阶段 = 7) AND ("触摸屏"."通风阶段运行时间（min）" <= 120));
   IF #_w1 THEN #催化加热温度上限 := "参数转换变量".M催化箱控制温度 + "参数转换变量".M催化箱控制温度上限; END_IF;
   "中间变量".催化加热控制阶段热回收阀打开 := #_w1;
   IF #_w1 THEN "中间变量".催化箱加热标志 := TRUE; END_IF;
   IF #_w1 AND ("触摸屏".催化前温度 <= "参数转换变量".M催化箱控制温度) THEN
       "中间变量".催化加热1标志 := TRUE;
       "中间变量".催化加热2标志 := TRUE;
   END_IF;
   IF #_w1 AND ("触摸屏".催化前温度 >= #催化加热温度上限) THEN
       "中间变量".催化加热1标志 := FALSE;
       "中间变量".催化加热2标志 := FALSE;
   END_IF;
   IF NOT "触摸屏".标志位1.%X1 AND NOT "触摸屏".手动操作1.%X0 THEN
       "中间变量".催化箱加热标志 := FALSE;
       "中间变量".催化加热1标志 := FALSE;
       "中间变量".催化加热2标志 := FALSE;
   END_IF;
END_REGION

REGION Network 2: 催化箱加热时间统计
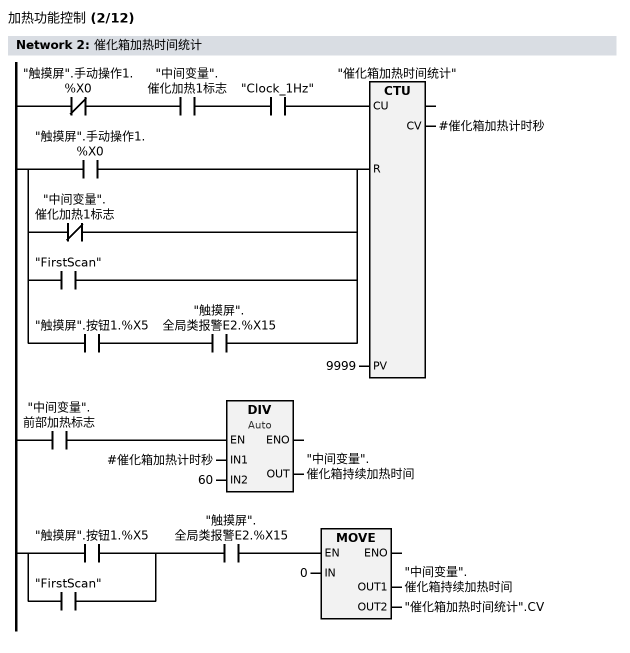
   "催化箱加热时间统计".CTU(CU := NOT "触摸屏".手动操作1.%X0 AND "中间变量".催化加热1标志 AND "Clock_1Hz",
                   R := "触摸屏".手动操作1.%X0 OR NOT "中间变量".催化加热1标志 OR "FirstScan" OR ("触摸屏".按钮1.%X5 AND "触摸屏".全局类报警E2.%X15),
                   PV := 9999,
                   CV => #催化箱加热计时秒);
   IF "中间变量".前部加热标志 THEN "中间变量".催化箱持续加热时间 := #催化箱加热计时秒 / 60; END_IF;
   IF ("触摸屏".按钮1.%X5 OR "FirstScan") AND "触摸屏".全局类报警E2.%X15 THEN
       "中间变量".催化箱持续加热时间 := 0;
       "催化箱加热时间统计".CV := 0;
   END_IF;
END_REGION

REGION Network 3: 汽化器温度加热控制
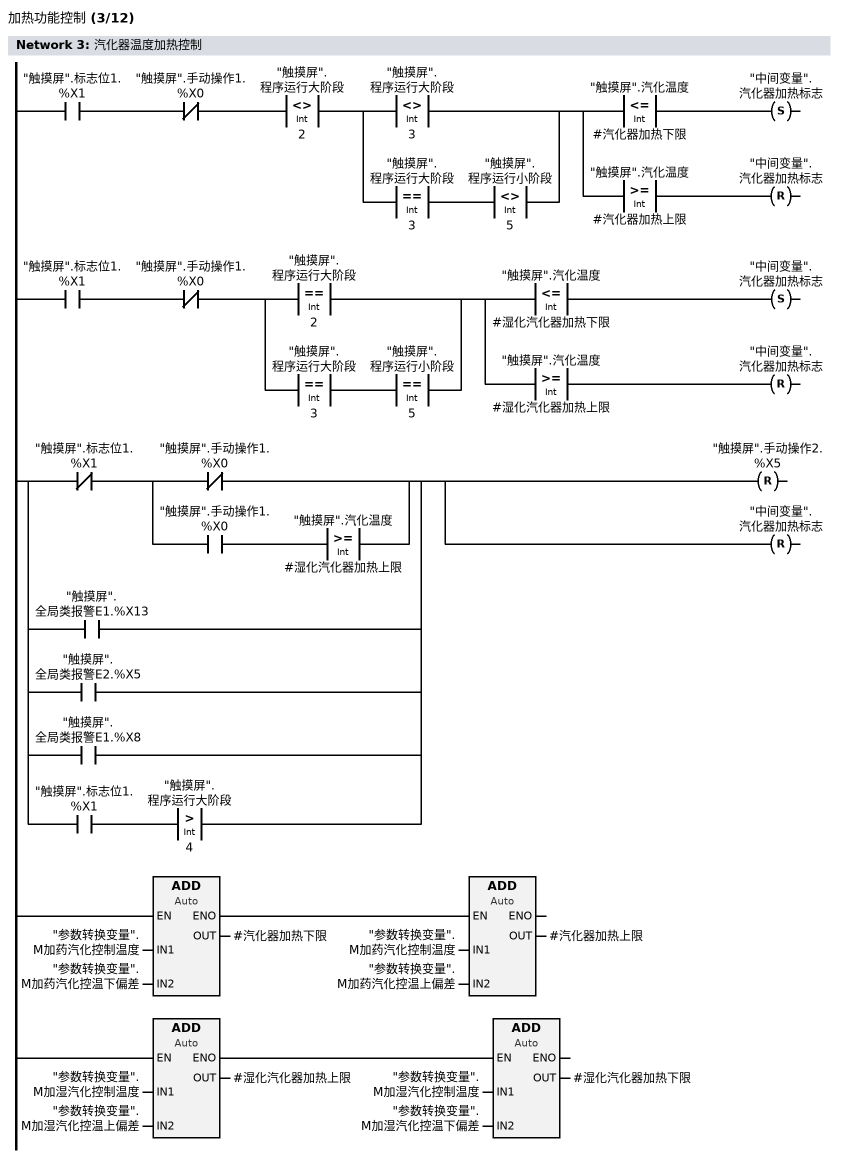
   RUNG wire#powerrail
      Contact( "触摸屏".标志位1.%X1 )
      I_Contact( "触摸屏".手动操作1.%X0 )
      { S7_Templates := "SrcType := Int" } NE_Contact(in1 := "触摸屏".程序运行大阶段, in2 := 2)
      wire#w1
      { S7_Templates := "SrcType := Int" } NE_Contact(in1 := "触摸屏".程序运行大阶段, in2 := 3)
      wire#w2
      { S7_Templates := "SrcType := Int" } LE_Contact(in1 := "触摸屏".汽化温度, in2 := #汽化器加热下限)
      S_Coil( "中间变量".汽化器加热标志 )
   END_RUNG
   RUNG wire#w1
      { S7_Templates := "SrcType := Int" } EQ_Contact(in1 := "触摸屏".程序运行大阶段, in2 := 3)
      { S7_Templates := "SrcType := Int" } NE_Contact(in1 := "触摸屏".程序运行小阶段, in2 := 5)
   END_RUNG wire#w2
   RUNG wire#w2
      { S7_Templates := "SrcType := Int" } GE_Contact(in1 := "触摸屏".汽化温度, in2 := #汽化器加热上限)
      R_Coil( "中间变量".汽化器加热标志 )
   END_RUNG
   RUNG wire#powerrail
      Contact( "触摸屏".标志位1.%X1 )
      I_Contact( "触摸屏".手动操作1.%X0 )
      wire#w3
      { S7_Templates := "SrcType := Int" } EQ_Contact(in1 := "触摸屏".程序运行大阶段, in2 := 2)
      wire#w4
      { S7_Templates := "SrcType := Int" } LE_Contact(in1 := "触摸屏".汽化温度, in2 := #湿化汽化器加热下限)
      S_Coil( "中间变量".汽化器加热标志 )
   END_RUNG
   RUNG wire#w3
      { S7_Templates := "SrcType := Int" } EQ_Contact(in1 := "触摸屏".程序运行大阶段, in2 := 3)
      { S7_Templates := "SrcType := Int" } EQ_Contact(in1 := "触摸屏".程序运行小阶段, in2 := 5)
   END_RUNG wire#w4
   RUNG wire#w4
      { S7_Templates := "SrcType := Int" } GE_Contact(in1 := "触摸屏".汽化温度, in2 := #湿化汽化器加热上限)
      R_Coil( "中间变量".汽化器加热标志 )
   END_RUNG
   RUNG wire#powerrail
      I_Contact( "触摸屏".标志位1.%X1 )
      wire#w5
      I_Contact( "触摸屏".手动操作1.%X0 )
      wire#w6
      R_Coil( "触摸屏".手动操作2.%X5 )
   END_RUNG
   RUNG wire#w5
      Contact( "触摸屏".手动操作1.%X0 )
      { S7_Templates := "SrcType := Int" } GE_Contact(in1 := "触摸屏".汽化温度, in2 := #湿化汽化器加热上限)
   END_RUNG wire#w6
   RUNG wire#powerrail
      Contact( "触摸屏".全局类报警E1.%X13 )
   END_RUNG wire#w6
   RUNG wire#powerrail
      Contact( "触摸屏".全局类报警E2.%X5 )
   END_RUNG wire#w6
   RUNG wire#powerrail
      Contact( "触摸屏".全局类报警E1.%X8 )
   END_RUNG wire#w6
   RUNG wire#powerrail
      Contact( "触摸屏".标志位1.%X1 )
      { S7_Templates := "SrcType := Int" } GT_Contact(in1 := "触摸屏".程序运行大阶段, in2 := 4)
   END_RUNG wire#w6
   RUNG wire#w6
      R_Coil( "中间变量".汽化器加热标志 )
   END_RUNG
   RUNG wire#powerrail
      Add(in1 := "参数转换变量".M加药汽化控制温度, in2 := "参数转换变量".M加药汽化控温下偏差, out => #汽化器加热下限)
      Add(in1 := "参数转换变量".M加药汽化控制温度, in2 := "参数转换变量".M加药汽化控温上偏差, out => #汽化器加热上限)
   END_RUNG
   RUNG wire#powerrail
      Add(in1 := "参数转换变量".M加湿汽化控制温度, in2 := "参数转换变量".M加湿汽化控温上偏差, out => #湿化汽化器加热上限)
      Add(in1 := "参数转换变量".M加湿汽化控制温度, in2 := "参数转换变量".M加湿汽化控温下偏差, out => #湿化汽化器加热下限)
   END_RUNG
   // the same network as SCL:
   #_w1 := "触摸屏".标志位1.%X1 AND NOT "触摸屏".手动操作1.%X0 AND ("触摸屏".程序运行大阶段 <> 2) AND (("触摸屏".程序运行大阶段 <> 3) OR (("触摸屏".程序运行大阶段 = 3) AND ("触摸屏".程序运行小阶段 <> 5)));
   IF #_w1 AND ("触摸屏".汽化温度 <= #汽化器加热下限) THEN "中间变量".汽化器加热标志 := TRUE; END_IF;
   IF #_w1 AND ("触摸屏".汽化温度 >= #汽化器加热上限) THEN "中间变量".汽化器加热标志 := FALSE; END_IF;
   #_w2 := "触摸屏".标志位1.%X1 AND NOT "触摸屏".手动操作1.%X0 AND (("触摸屏".程序运行大阶段 = 2) OR (("触摸屏".程序运行大阶段 = 3) AND ("触摸屏".程序运行小阶段 = 5)));
   IF #_w2 AND ("触摸屏".汽化温度 <= #湿化汽化器加热下限) THEN "中间变量".汽化器加热标志 := TRUE; END_IF;
   IF #_w2 AND ("触摸屏".汽化温度 >= #湿化汽化器加热上限) THEN "中间变量".汽化器加热标志 := FALSE; END_IF;
   IF (NOT "触摸屏".标志位1.%X1 AND (NOT "触摸屏".手动操作1.%X0 OR ("触摸屏".手动操作1.%X0 AND ("触摸屏".汽化温度 >= #湿化汽化器加热上限)))) OR "触摸屏".全局类报警E1.%X13 OR "触摸屏".全局类报警E2.%X5 OR "触摸屏".全局类报警E1.%X8 OR ("触摸屏".标志位1.%X1 AND ("触摸屏".程序运行大阶段 > 4)) THEN
       "触摸屏".手动操作2.%X5 := FALSE;
       "中间变量".汽化器加热标志 := FALSE;
   END_IF;
   #汽化器加热下限 := "参数转换变量".M加药汽化控制温度 + "参数转换变量".M加药汽化控温下偏差;
   #汽化器加热上限 := "参数转换变量".M加药汽化控制温度 + "参数转换变量".M加药汽化控温上偏差;
   #湿化汽化器加热上限 := "参数转换变量".M加湿汽化控制温度 + "参数转换变量".M加湿汽化控温上偏差;
   #湿化汽化器加热下限 := "参数转换变量".M加湿汽化控制温度 + "参数转换变量".M加湿汽化控温下偏差;
END_REGION

REGION Network 4: 汽化器温度加热控制时间统计
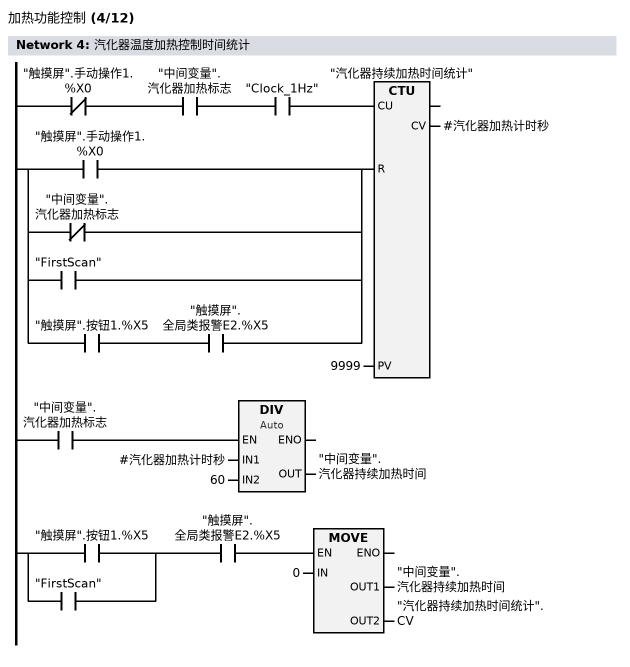
   "汽化器持续加热时间统计".CTU(CU := NOT "触摸屏".手动操作1.%X0 AND "中间变量".汽化器加热标志 AND "Clock_1Hz",
                     R := "触摸屏".手动操作1.%X0 OR NOT "中间变量".汽化器加热标志 OR "FirstScan" OR ("触摸屏".按钮1.%X5 AND "触摸屏".全局类报警E2.%X5),
                     PV := 9999,
                     CV => #汽化器加热计时秒);
   IF "中间变量".汽化器加热标志 THEN "中间变量".汽化器持续加热时间 := #汽化器加热计时秒 / 60; END_IF;
   IF ("触摸屏".按钮1.%X5 OR "FirstScan") AND "触摸屏".全局类报警E2.%X5 THEN
       "中间变量".汽化器持续加热时间 := 0;
       "汽化器持续加热时间统计".CV := 0;
   END_IF;
END_REGION

REGION Network 5: 腔体前部加热
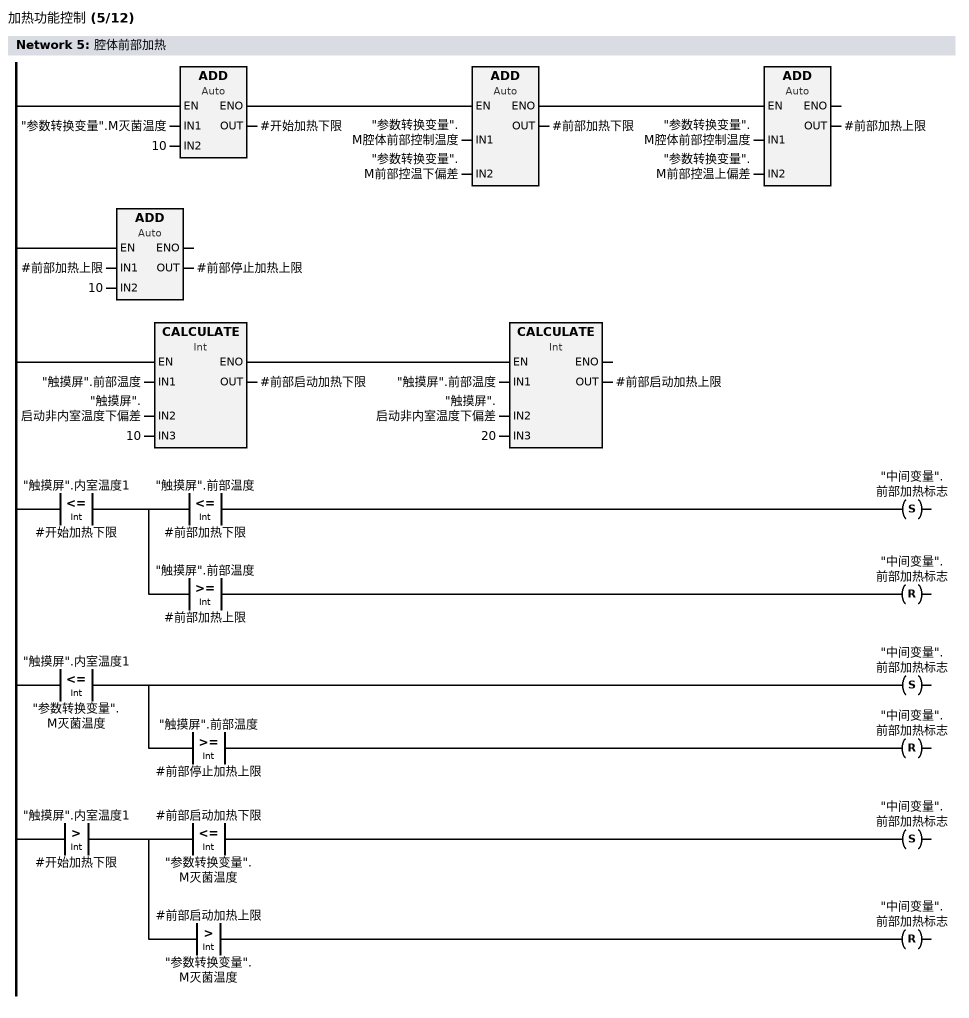
   RUNG wire#powerrail
      Add(in1 := "参数转换变量".M灭菌温度, in2 := 10, out => #开始加热下限)
      Add(in1 := "参数转换变量".M腔体前部控制温度, in2 := "参数转换变量".M前部控温下偏差, out => #前部加热下限)
      Add(in1 := "参数转换变量".M腔体前部控制温度, in2 := "参数转换变量".M前部控温上偏差, out => #前部加热上限)
   END_RUNG
   RUNG wire#powerrail
      Add(in1 := #前部加热上限, in2 := 10, out => #前部停止加热上限)
   END_RUNG
   RUNG wire#powerrail
      { S7_Templates := "SrcType := Int"; S7_Expression := "IN1+IN2-IN3" } Calculate(in1 := "触摸屏".前部温度, in2 := "触摸屏".启动非内室温度下偏差, in3 := 10, out => #前部启动加热下限)
      { S7_Templates := "SrcType := Int"; S7_Expression := "IN1+IN2-IN3" } Calculate(in1 := "触摸屏".前部温度, in2 := "触摸屏".启动非内室温度下偏差, in3 := 20, out => #前部启动加热上限)
   END_RUNG
   RUNG wire#powerrail
      { S7_Templates := "SrcType := Int" } LE_Contact(in1 := "触摸屏".内室温度1, in2 := #开始加热下限)
      wire#w1
      { S7_Templates := "SrcType := Int" } LE_Contact(in1 := "触摸屏".前部温度, in2 := #前部加热下限)
      S_Coil( "中间变量".前部加热标志 )
   END_RUNG
   RUNG wire#w1
      { S7_Templates := "SrcType := Int" } GE_Contact(in1 := "触摸屏".前部温度, in2 := #前部加热上限)
      R_Coil( "中间变量".前部加热标志 )
   END_RUNG
   RUNG wire#powerrail
      { S7_Templates := "SrcType := Int" } LE_Contact(in1 := "触摸屏".内室温度1, in2 := "参数转换变量".M灭菌温度)
      wire#w2
      S_Coil( "中间变量".前部加热标志 )
   END_RUNG
   RUNG wire#w2
      { S7_Templates := "SrcType := Int" } GE_Contact(in1 := "触摸屏".前部温度, in2 := #前部停止加热上限)
      R_Coil( "中间变量".前部加热标志 )
   END_RUNG
   RUNG wire#powerrail
      { S7_Templates := "SrcType := Int" } GT_Contact(in1 := "触摸屏".内室温度1, in2 := #开始加热下限)
      wire#w3
      { S7_Templates := "SrcType := Int" } LE_Contact(in1 := #前部启动加热下限, in2 := "参数转换变量".M灭菌温度)
      S_Coil( "中间变量".前部加热标志 )
   END_RUNG
   RUNG wire#w3
      { S7_Templates := "SrcType := Int" } GT_Contact(in1 := #前部启动加热上限, in2 := "参数转换变量".M灭菌温度)
      R_Coil( "中间变量".前部加热标志 )
   END_RUNG
   // the same network as SCL:
   #开始加热下限 := "参数转换变量".M灭菌温度 + 10;
   #前部加热下限 := "参数转换变量".M腔体前部控制温度 + "参数转换变量".M前部控温下偏差;
   #前部加热上限 := "参数转换变量".M腔体前部控制温度 + "参数转换变量".M前部控温上偏差;
   #前部停止加热上限 := #前部加热上限 + 10;
   #前部启动加热下限 := "触摸屏".前部温度+"触摸屏".启动非内室温度下偏差-10;
   #前部启动加热上限 := "触摸屏".前部温度+"触摸屏".启动非内室温度下偏差-20;
   #_w1 := "触摸屏".内室温度1 <= #开始加热下限;
   IF #_w1 AND ("触摸屏".前部温度 <= #前部加热下限) THEN "中间变量".前部加热标志 := TRUE; END_IF;
   IF #_w1 AND ("触摸屏".前部温度 >= #前部加热上限) THEN "中间变量".前部加热标志 := FALSE; END_IF;
   #_w2 := "触摸屏".内室温度1 <= "参数转换变量".M灭菌温度;
   IF #_w2 THEN "中间变量".前部加热标志 := TRUE; END_IF;
   IF #_w2 AND ("触摸屏".前部温度 >= #前部停止加热上限) THEN "中间变量".前部加热标志 := FALSE; END_IF;
   #_w3 := "触摸屏".内室温度1 > #开始加热下限;
   IF #_w3 AND (#前部启动加热下限 <= "参数转换变量".M灭菌温度) THEN "中间变量".前部加热标志 := TRUE; END_IF;
   IF #_w3 AND (#前部启动加热上限 > "参数转换变量".M灭菌温度) THEN "中间变量".前部加热标志 := FALSE; END_IF;
END_REGION

REGION Network 6: 腔体前部加热时间统计
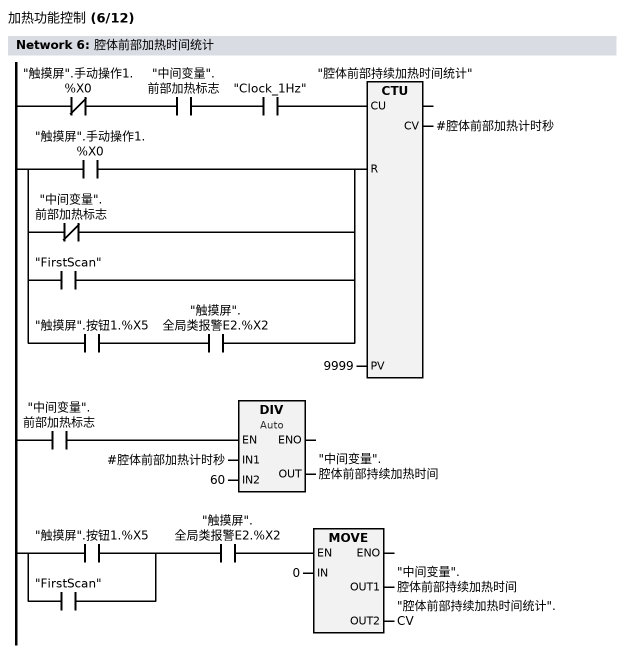
   "腔体前部持续加热时间统计".CTU(CU := NOT "触摸屏".手动操作1.%X0 AND "中间变量".前部加热标志 AND "Clock_1Hz",
                      R := "触摸屏".手动操作1.%X0 OR NOT "中间变量".前部加热标志 OR "FirstScan" OR ("触摸屏".按钮1.%X5 AND "触摸屏".全局类报警E2.%X2),
                      PV := 9999,
                      CV => #腔体前部加热计时秒);
   IF "中间变量".前部加热标志 THEN "中间变量".腔体前部持续加热时间 := #腔体前部加热计时秒 / 60; END_IF;
   IF ("触摸屏".按钮1.%X5 OR "FirstScan") AND "触摸屏".全局类报警E2.%X2 THEN
       "中间变量".腔体前部持续加热时间 := 0;
       "腔体前部持续加热时间统计".CV := 0;
   END_IF;
END_REGION

REGION Network 7: 腔体后部加热
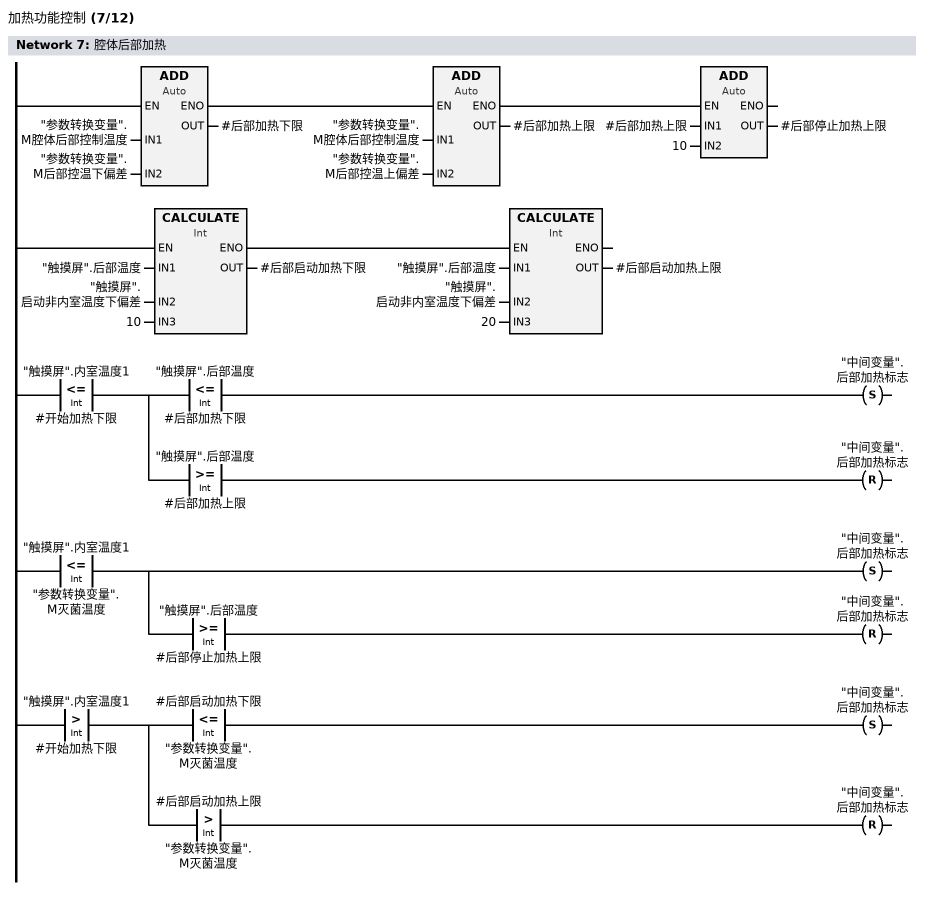
   RUNG wire#powerrail
      Add(in1 := "参数转换变量".M腔体后部控制温度, in2 := "参数转换变量".M后部控温下偏差, out => #后部加热下限)
      Add(in1 := "参数转换变量".M腔体后部控制温度, in2 := "参数转换变量".M后部控温上偏差, out => #后部加热上限)
      Add(in1 := #后部加热上限, in2 := 10, out => #后部停止加热上限)
   END_RUNG
   RUNG wire#powerrail
      { S7_Templates := "SrcType := Int"; S7_Expression := "IN1+IN2-IN3" } Calculate(in1 := "触摸屏".后部温度, in2 := "触摸屏".启动非内室温度下偏差, in3 := 10, out => #后部启动加热下限)
      { S7_Templates := "SrcType := Int"; S7_Expression := "IN1+IN2-IN3" } Calculate(in1 := "触摸屏".后部温度, in2 := "触摸屏".启动非内室温度下偏差, in3 := 20, out => #后部启动加热上限)
   END_RUNG
   RUNG wire#powerrail
      { S7_Templates := "SrcType := Int" } LE_Contact(in1 := "触摸屏".内室温度1, in2 := #开始加热下限)
      wire#w1
      { S7_Templates := "SrcType := Int" } LE_Contact(in1 := "触摸屏".后部温度, in2 := #后部加热下限)
      S_Coil( "中间变量".后部加热标志 )
   END_RUNG
   RUNG wire#w1
      { S7_Templates := "SrcType := Int" } GE_Contact(in1 := "触摸屏".后部温度, in2 := #后部加热上限)
      R_Coil( "中间变量".后部加热标志 )
   END_RUNG
   RUNG wire#powerrail
      { S7_Templates := "SrcType := Int" } LE_Contact(in1 := "触摸屏".内室温度1, in2 := "参数转换变量".M灭菌温度)
      wire#w2
      S_Coil( "中间变量".后部加热标志 )
   END_RUNG
   RUNG wire#w2
      { S7_Templates := "SrcType := Int" } GE_Contact(in1 := "触摸屏".后部温度, in2 := #后部停止加热上限)
      R_Coil( "中间变量".后部加热标志 )
   END_RUNG
   RUNG wire#powerrail
      { S7_Templates := "SrcType := Int" } GT_Contact(in1 := "触摸屏".内室温度1, in2 := #开始加热下限)
      wire#w3
      { S7_Templates := "SrcType := Int" } LE_Contact(in1 := #后部启动加热下限, in2 := "参数转换变量".M灭菌温度)
      S_Coil( "中间变量".后部加热标志 )
   END_RUNG
   RUNG wire#w3
      { S7_Templates := "SrcType := Int" } GT_Contact(in1 := #后部启动加热上限, in2 := "参数转换变量".M灭菌温度)
      R_Coil( "中间变量".后部加热标志 )
   END_RUNG
   // the same network as SCL:
   #后部加热下限 := "参数转换变量".M腔体后部控制温度 + "参数转换变量".M后部控温下偏差;
   #后部加热上限 := "参数转换变量".M腔体后部控制温度 + "参数转换变量".M后部控温上偏差;
   #后部停止加热上限 := #后部加热上限 + 10;
   #后部启动加热下限 := "触摸屏".后部温度+"触摸屏".启动非内室温度下偏差-10;
   #后部启动加热上限 := "触摸屏".后部温度+"触摸屏".启动非内室温度下偏差-20;
   #_w1 := "触摸屏".内室温度1 <= #开始加热下限;
   IF #_w1 AND ("触摸屏".后部温度 <= #后部加热下限) THEN "中间变量".后部加热标志 := TRUE; END_IF;
   IF #_w1 AND ("触摸屏".后部温度 >= #后部加热上限) THEN "中间变量".后部加热标志 := FALSE; END_IF;
   #_w2 := "触摸屏".内室温度1 <= "参数转换变量".M灭菌温度;
   IF #_w2 THEN "中间变量".后部加热标志 := TRUE; END_IF;
   IF #_w2 AND ("触摸屏".后部温度 >= #后部停止加热上限) THEN "中间变量".后部加热标志 := FALSE; END_IF;
   #_w3 := "触摸屏".内室温度1 > #开始加热下限;
   IF #_w3 AND (#后部启动加热下限 <= "参数转换变量".M灭菌温度) THEN "中间变量".后部加热标志 := TRUE; END_IF;
   IF #_w3 AND (#后部启动加热上限 > "参数转换变量".M灭菌温度) THEN "中间变量".后部加热标志 := FALSE; END_IF;
END_REGION

REGION Network 8: 腔体后部加热时间统计
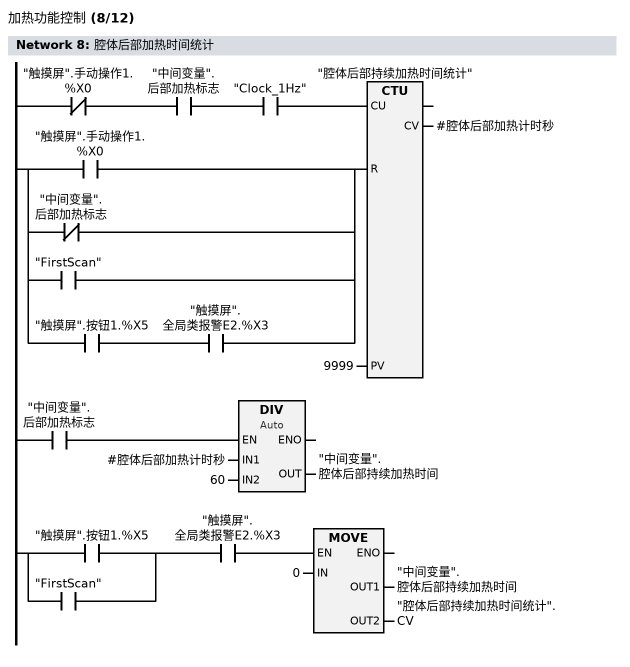
   "腔体后部持续加热时间统计".CTU(CU := NOT "触摸屏".手动操作1.%X0 AND "中间变量".后部加热标志 AND "Clock_1Hz",
                      R := "触摸屏".手动操作1.%X0 OR NOT "中间变量".后部加热标志 OR "FirstScan" OR ("触摸屏".按钮1.%X5 AND "触摸屏".全局类报警E2.%X3),
                      PV := 9999,
                      CV => #腔体后部加热计时秒);
   IF "中间变量".后部加热标志 THEN "中间变量".腔体后部持续加热时间 := #腔体后部加热计时秒 / 60; END_IF;
   IF ("触摸屏".按钮1.%X5 OR "FirstScan") AND "触摸屏".全局类报警E2.%X3 THEN
       "中间变量".腔体后部持续加热时间 := 0;
       "腔体后部持续加热时间统计".CV := 0;
   END_IF;
END_REGION

REGION Network 9: 前门加热
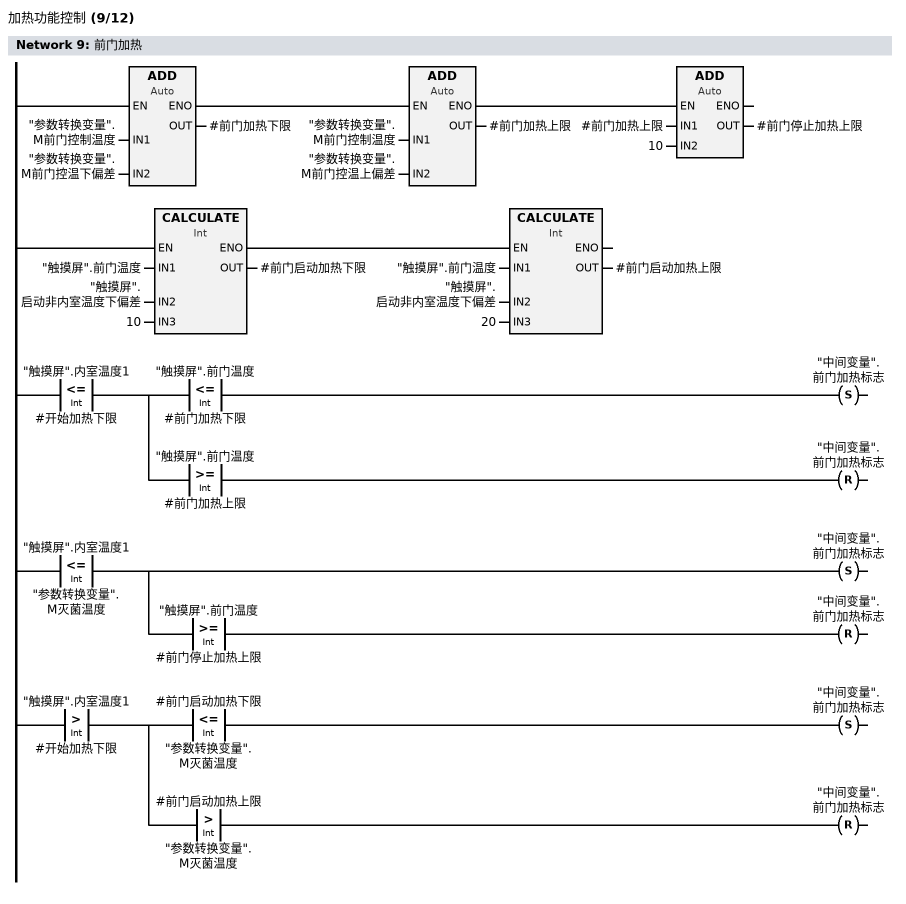
   RUNG wire#powerrail
      Add(in1 := "参数转换变量".M前门控制温度, in2 := "参数转换变量".M前门控温下偏差, out => #前门加热下限)
      Add(in1 := "参数转换变量".M前门控制温度, in2 := "参数转换变量".M前门控温上偏差, out => #前门加热上限)
      Add(in1 := #前门加热上限, in2 := 10, out => #前门停止加热上限)
   END_RUNG
   RUNG wire#powerrail
      { S7_Templates := "SrcType := Int"; S7_Expression := "IN1+IN2-IN3" } Calculate(in1 := "触摸屏".前门温度, in2 := "触摸屏".启动非内室温度下偏差, in3 := 10, out => #前门启动加热下限)
      { S7_Templates := "SrcType := Int"; S7_Expression := "IN1+IN2-IN3" } Calculate(in1 := "触摸屏".前门温度, in2 := "触摸屏".启动非内室温度下偏差, in3 := 20, out => #前门启动加热上限)
   END_RUNG
   RUNG wire#powerrail
      { S7_Templates := "SrcType := Int" } LE_Contact(in1 := "触摸屏".内室温度1, in2 := #开始加热下限)
      wire#w1
      { S7_Templates := "SrcType := Int" } LE_Contact(in1 := "触摸屏".前门温度, in2 := #前门加热下限)
      S_Coil( "中间变量".前门加热标志 )
   END_RUNG
   RUNG wire#w1
      { S7_Templates := "SrcType := Int" } GE_Contact(in1 := "触摸屏".前门温度, in2 := #前门加热上限)
      R_Coil( "中间变量".前门加热标志 )
   END_RUNG
   RUNG wire#powerrail
      { S7_Templates := "SrcType := Int" } LE_Contact(in1 := "触摸屏".内室温度1, in2 := "参数转换变量".M灭菌温度)
      wire#w2
      S_Coil( "中间变量".前门加热标志 )
   END_RUNG
   RUNG wire#w2
      { S7_Templates := "SrcType := Int" } GE_Contact(in1 := "触摸屏".前门温度, in2 := #前门停止加热上限)
      R_Coil( "中间变量".前门加热标志 )
   END_RUNG
   RUNG wire#powerrail
      { S7_Templates := "SrcType := Int" } GT_Contact(in1 := "触摸屏".内室温度1, in2 := #开始加热下限)
      wire#w3
      { S7_Templates := "SrcType := Int" } LE_Contact(in1 := #前门启动加热下限, in2 := "参数转换变量".M灭菌温度)
      S_Coil( "中间变量".前门加热标志 )
   END_RUNG
   RUNG wire#w3
      { S7_Templates := "SrcType := Int" } GT_Contact(in1 := #前门启动加热上限, in2 := "参数转换变量".M灭菌温度)
      R_Coil( "中间变量".前门加热标志 )
   END_RUNG
   // the same network as SCL:
   #前门加热下限 := "参数转换变量".M前门控制温度 + "参数转换变量".M前门控温下偏差;
   #前门加热上限 := "参数转换变量".M前门控制温度 + "参数转换变量".M前门控温上偏差;
   #前门停止加热上限 := #前门加热上限 + 10;
   #前门启动加热下限 := "触摸屏".前门温度+"触摸屏".启动非内室温度下偏差-10;
   #前门启动加热上限 := "触摸屏".前门温度+"触摸屏".启动非内室温度下偏差-20;
   #_w1 := "触摸屏".内室温度1 <= #开始加热下限;
   IF #_w1 AND ("触摸屏".前门温度 <= #前门加热下限) THEN "中间变量".前门加热标志 := TRUE; END_IF;
   IF #_w1 AND ("触摸屏".前门温度 >= #前门加热上限) THEN "中间变量".前门加热标志 := FALSE; END_IF;
   #_w2 := "触摸屏".内室温度1 <= "参数转换变量".M灭菌温度;
   IF #_w2 THEN "中间变量".前门加热标志 := TRUE; END_IF;
   IF #_w2 AND ("触摸屏".前门温度 >= #前门停止加热上限) THEN "中间变量".前门加热标志 := FALSE; END_IF;
   #_w3 := "触摸屏".内室温度1 > #开始加热下限;
   IF #_w3 AND (#前门启动加热下限 <= "参数转换变量".M灭菌温度) THEN "中间变量".前门加热标志 := TRUE; END_IF;
   IF #_w3 AND (#前门启动加热上限 > "参数转换变量".M灭菌温度) THEN "中间变量".前门加热标志 := FALSE; END_IF;
END_REGION

REGION Network 10: 前门加热时间统计
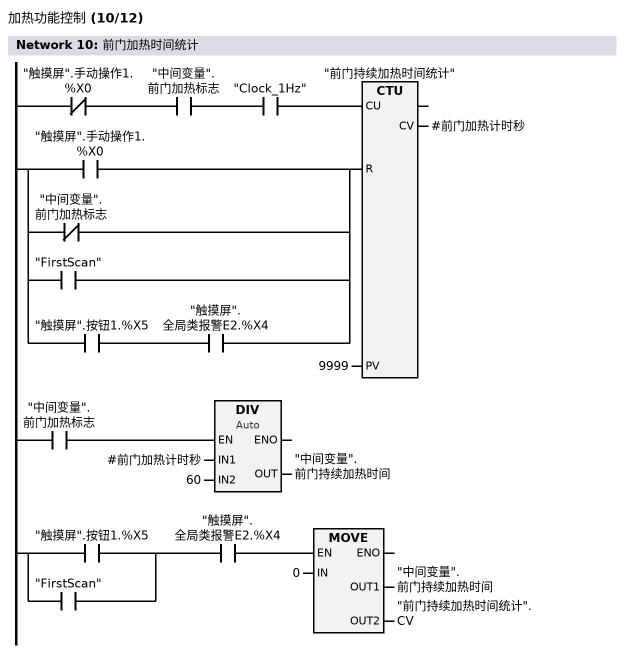
   "前门持续加热时间统计".CTU(CU := NOT "触摸屏".手动操作1.%X0 AND "中间变量".前门加热标志 AND "Clock_1Hz",
                    R := "触摸屏".手动操作1.%X0 OR NOT "中间变量".前门加热标志 OR "FirstScan" OR ("触摸屏".按钮1.%X5 AND "触摸屏".全局类报警E2.%X4),
                    PV := 9999,
                    CV => #前门加热计时秒);
   IF "中间变量".前门加热标志 THEN "中间变量".前门持续加热时间 := #前门加热计时秒 / 60; END_IF;
   IF ("触摸屏".按钮1.%X5 OR "FirstScan") AND "触摸屏".全局类报警E2.%X4 THEN
       "中间变量".前门持续加热时间 := 0;
       "前门持续加热时间统计".CV := 0;
   END_IF;
END_REGION

REGION Network 11: 后门加热
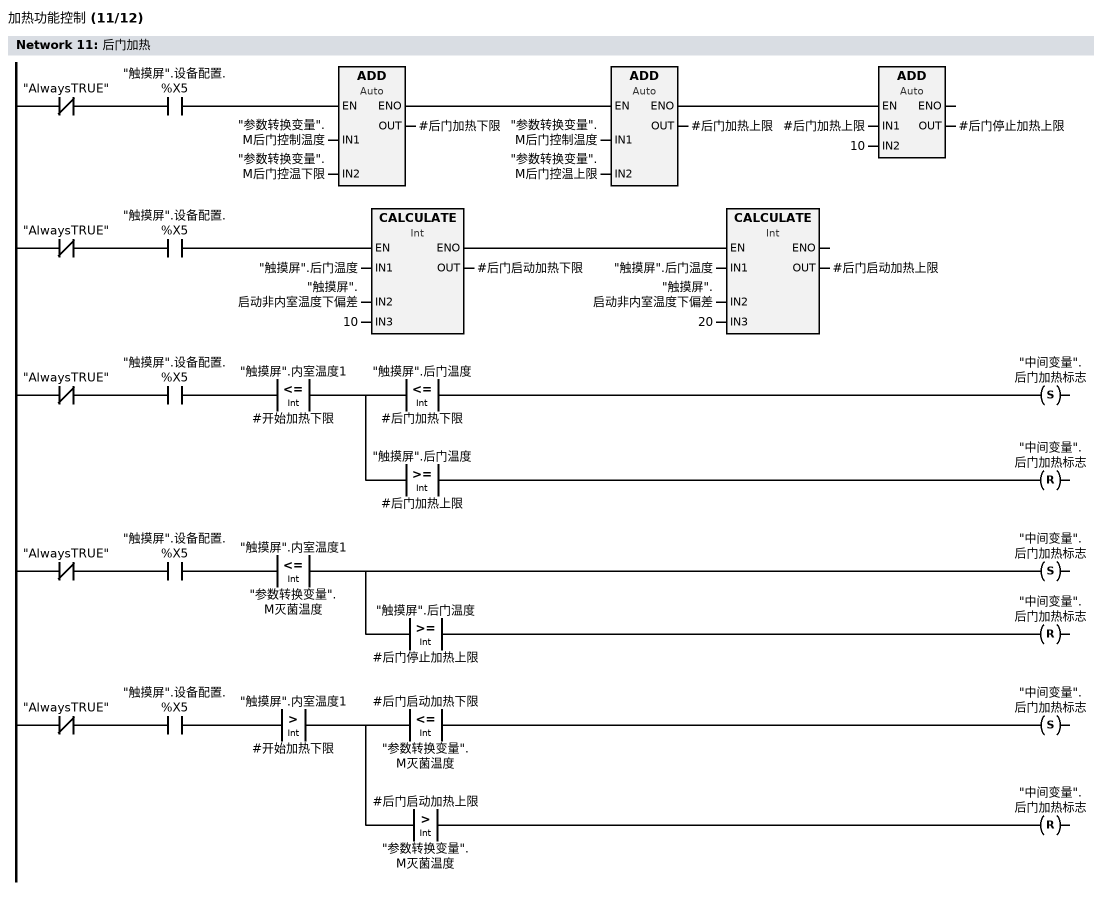
   RUNG wire#powerrail
      I_Contact( "AlwaysTRUE" )
      Contact( "触摸屏".设备配置.%X5 )
      Add(in1 := "参数转换变量".M后门控制温度, in2 := "参数转换变量".M后门控温下限, out => #后门加热下限)
      Add(in1 := "参数转换变量".M后门控制温度, in2 := "参数转换变量".M后门控温上限, out => #后门加热上限)
      Add(in1 := #后门加热上限, in2 := 10, out => #后门停止加热上限)
   END_RUNG
   RUNG wire#powerrail
      I_Contact( "AlwaysTRUE" )
      Contact( "触摸屏".设备配置.%X5 )
      { S7_Templates := "SrcType := Int"; S7_Expression := "IN1+IN2-IN3" } Calculate(in1 := "触摸屏".后门温度, in2 := "触摸屏".启动非内室温度下偏差, in3 := 10, out => #后门启动加热下限)
      { S7_Templates := "SrcType := Int"; S7_Expression := "IN1+IN2-IN3" } Calculate(in1 := "触摸屏".后门温度, in2 := "触摸屏".启动非内室温度下偏差, in3 := 20, out => #后门启动加热上限)
   END_RUNG
   RUNG wire#powerrail
      I_Contact( "AlwaysTRUE" )
      Contact( "触摸屏".设备配置.%X5 )
      { S7_Templates := "SrcType := Int" } LE_Contact(in1 := "触摸屏".内室温度1, in2 := #开始加热下限)
      wire#w1
      { S7_Templates := "SrcType := Int" } LE_Contact(in1 := "触摸屏".后门温度, in2 := #后门加热下限)
      S_Coil( "中间变量".后门加热标志 )
   END_RUNG
   RUNG wire#w1
      { S7_Templates := "SrcType := Int" } GE_Contact(in1 := "触摸屏".后门温度, in2 := #后门加热上限)
      R_Coil( "中间变量".后门加热标志 )
   END_RUNG
   RUNG wire#powerrail
      I_Contact( "AlwaysTRUE" )
      Contact( "触摸屏".设备配置.%X5 )
      { S7_Templates := "SrcType := Int" } LE_Contact(in1 := "触摸屏".内室温度1, in2 := "参数转换变量".M灭菌温度)
      wire#w2
      S_Coil( "中间变量".后门加热标志 )
   END_RUNG
   RUNG wire#w2
      { S7_Templates := "SrcType := Int" } GE_Contact(in1 := "触摸屏".后门温度, in2 := #后门停止加热上限)
      R_Coil( "中间变量".后门加热标志 )
   END_RUNG
   RUNG wire#powerrail
      I_Contact( "AlwaysTRUE" )
      Contact( "触摸屏".设备配置.%X5 )
      { S7_Templates := "SrcType := Int" } GT_Contact(in1 := "触摸屏".内室温度1, in2 := #开始加热下限)
      wire#w3
      { S7_Templates := "SrcType := Int" } LE_Contact(in1 := #后门启动加热下限, in2 := "参数转换变量".M灭菌温度)
      S_Coil( "中间变量".后门加热标志 )
   END_RUNG
   RUNG wire#w3
      { S7_Templates := "SrcType := Int" } GT_Contact(in1 := #后门启动加热上限, in2 := "参数转换变量".M灭菌温度)
      R_Coil( "中间变量".后门加热标志 )
   END_RUNG
   // the same network as SCL:
   IF NOT "AlwaysTRUE" AND "触摸屏".设备配置.%X5 THEN
       #后门加热下限 := "参数转换变量".M后门控制温度 + "参数转换变量".M后门控温下限;
       #后门加热上限 := "参数转换变量".M后门控制温度 + "参数转换变量".M后门控温上限;
       #后门停止加热上限 := #后门加热上限 + 10;
       #后门启动加热下限 := "触摸屏".后门温度+"触摸屏".启动非内室温度下偏差-10;
       #后门启动加热上限 := "触摸屏".后门温度+"触摸屏".启动非内室温度下偏差-20;
   END_IF;
   #_w1 := NOT "AlwaysTRUE" AND "触摸屏".设备配置.%X5 AND ("触摸屏".内室温度1 <= #开始加热下限);
   IF #_w1 AND ("触摸屏".后门温度 <= #后门加热下限) THEN "中间变量".后门加热标志 := TRUE; END_IF;
   IF #_w1 AND ("触摸屏".后门温度 >= #后门加热上限) THEN "中间变量".后门加热标志 := FALSE; END_IF;
   #_w2 := NOT "AlwaysTRUE" AND "触摸屏".设备配置.%X5 AND ("触摸屏".内室温度1 <= "参数转换变量".M灭菌温度);
   IF #_w2 THEN "中间变量".后门加热标志 := TRUE; END_IF;
   IF #_w2 AND ("触摸屏".后门温度 >= #后门停止加热上限) THEN "中间变量".后门加热标志 := FALSE; END_IF;
   #_w3 := NOT "AlwaysTRUE" AND "触摸屏".设备配置.%X5 AND ("触摸屏".内室温度1 > #开始加热下限);
   IF #_w3 AND (#后门启动加热下限 <= "参数转换变量".M灭菌温度) THEN "中间变量".后门加热标志 := TRUE; END_IF;
   IF #_w3 AND (#后门启动加热上限 > "参数转换变量".M灭菌温度) THEN "中间变量".后门加热标志 := FALSE; END_IF;
END_REGION

REGION Network 12: 后门加热时间统计
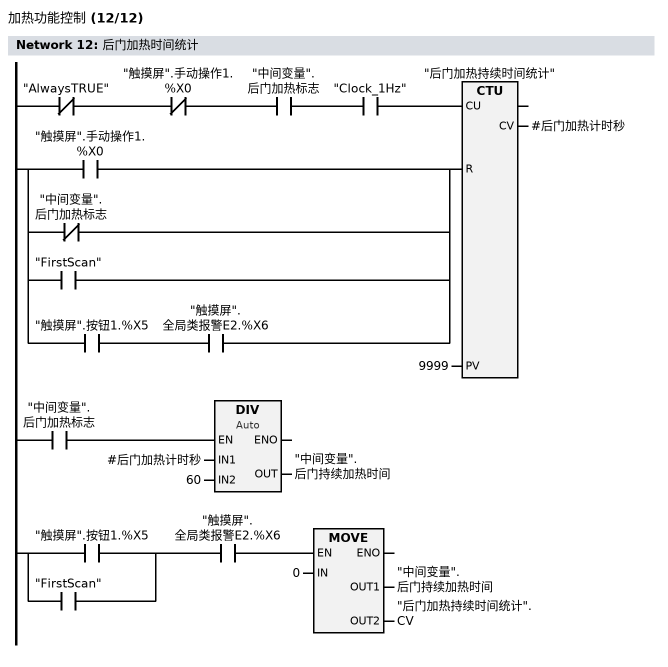
   "后门加热持续时间统计".CTU(CU := NOT "AlwaysTRUE" AND NOT "触摸屏".手动操作1.%X0 AND "中间变量".后门加热标志 AND "Clock_1Hz",
                    R := "触摸屏".手动操作1.%X0 OR NOT "中间变量".后门加热标志 OR "FirstScan" OR ("触摸屏".按钮1.%X5 AND "触摸屏".全局类报警E2.%X6),
                    PV := 9999,
                    CV => #后门加热计时秒);
   IF "中间变量".后门加热标志 THEN "中间变量".后门持续加热时间 := #后门加热计时秒 / 60; END_IF;
   IF ("触摸屏".按钮1.%X5 OR "FirstScan") AND "触摸屏".全局类报警E2.%X6 THEN
       "中间变量".后门持续加热时间 := 0;
       "后门加热持续时间统计".CV := 0;
   END_IF;
END_REGION
END_FUNCTION_BLOCK

// folder: 16数字量输出

FUNCTION "数字量输出控制" : Void   // FC5, LAD
{ S7_Optimized_Access := 'TRUE' }
VERSION : 0.1
BEGIN

REGION Network 1: 回空阀V1
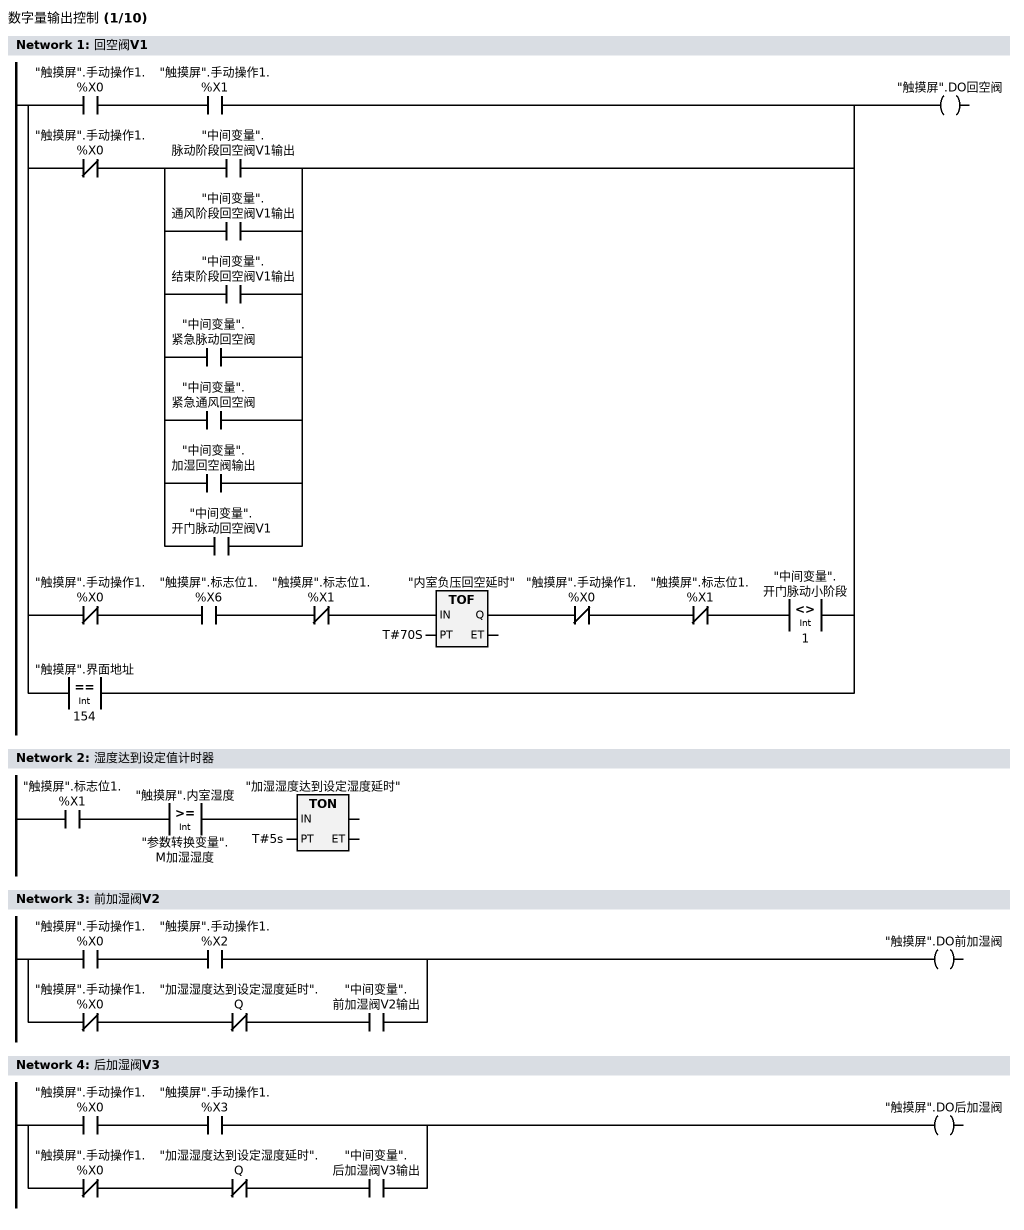
   "内室负压回空延时".TOF(IN := NOT "触摸屏".手动操作1.%X0 AND "触摸屏".标志位1.%X6 AND NOT "触摸屏".标志位1.%X1, PT := T#70S);
   "触摸屏".DO回空阀 := ("触摸屏".手动操作1.%X0 AND "触摸屏".手动操作1.%X1) OR (NOT "触摸屏".手动操作1.%X0 AND ("中间变量".脉动阶段回空阀V1输出 OR "中间变量".通风阶段回空阀V1输出 OR "中间变量".结束阶段回空阀V1输出 OR "中间变量".紧急脉动回空阀 OR "中间变量".紧急通风回空阀 OR "中间变量".加湿回空阀输出 OR "中间变量".开门脉动回空阀V1)) OR ("内室负压回空延时".Q AND NOT "触摸屏".手动操作1.%X0 AND NOT "触摸屏".标志位1.%X1 AND ("中间变量".开门脉动小阶段 <> 1)) OR ("触摸屏".界面地址 = 154);
END_REGION

REGION Network 2: 湿度达到设定值计时器
   "加湿湿度达到设定湿度延时".TON(IN := "触摸屏".标志位1.%X1 AND ("触摸屏".内室湿度 >= "参数转换变量".M加湿湿度), PT := T#5s);
END_REGION

REGION Network 3: 前加湿阀V2
   RUNG wire#powerrail
      Contact( "触摸屏".手动操作1.%X0 )
      Contact( "触摸屏".手动操作1.%X2 )
      wire#w1
      Coil( "触摸屏".DO前加湿阀 )
   END_RUNG
   RUNG wire#powerrail
      I_Contact( "触摸屏".手动操作1.%X0 )
      I_Contact( "加湿湿度达到设定湿度延时".Q )
      Contact( "中间变量".前加湿阀V2输出 )
   END_RUNG wire#w1
   // the same network as SCL:
   "触摸屏".DO前加湿阀 := ("触摸屏".手动操作1.%X0 AND "触摸屏".手动操作1.%X2) OR (NOT "触摸屏".手动操作1.%X0 AND NOT "加湿湿度达到设定湿度延时".Q AND "中间变量".前加湿阀V2输出);
END_REGION

REGION Network 4: 后加湿阀V3
   RUNG wire#powerrail
      Contact( "触摸屏".手动操作1.%X0 )
      Contact( "触摸屏".手动操作1.%X3 )
      wire#w1
      Coil( "触摸屏".DO后加湿阀 )
   END_RUNG
   RUNG wire#powerrail
      I_Contact( "触摸屏".手动操作1.%X0 )
      I_Contact( "加湿湿度达到设定湿度延时".Q )
      Contact( "中间变量".后加湿阀V3输出 )
   END_RUNG wire#w1
   // the same network as SCL:
   "触摸屏".DO后加湿阀 := ("触摸屏".手动操作1.%X0 AND "触摸屏".手动操作1.%X3) OR (NOT "触摸屏".手动操作1.%X0 AND NOT "加湿湿度达到设定湿度延时".Q AND "中间变量".后加湿阀V3输出);
END_REGION

REGION Network 5: 快抽空阀V4
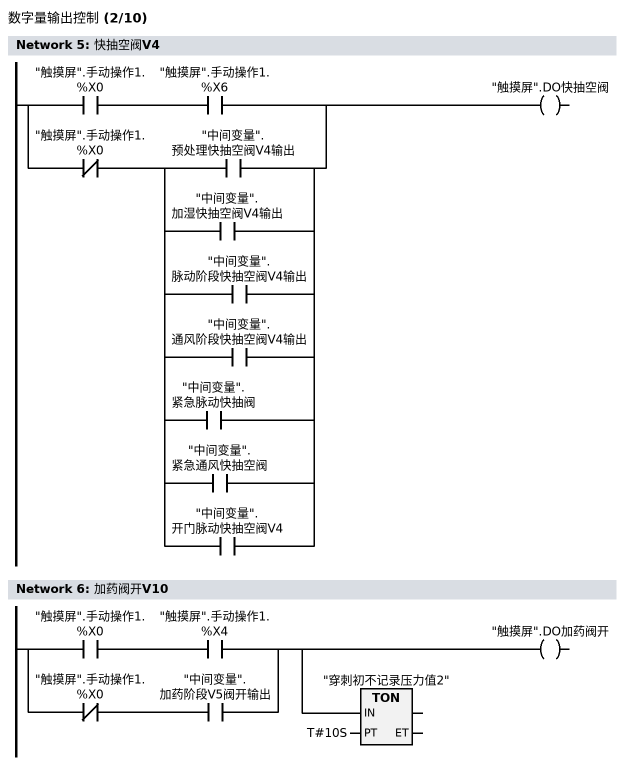
   RUNG wire#powerrail
      Contact( "触摸屏".手动操作1.%X0 )
      Contact( "触摸屏".手动操作1.%X6 )
      wire#w1
      Coil( "触摸屏".DO快抽空阀 )
   END_RUNG
   RUNG wire#powerrail
      I_Contact( "触摸屏".手动操作1.%X0 )
      wire#w2
      Contact( "中间变量".预处理快抽空阀V4输出 )
   END_RUNG wire#w1
   RUNG wire#w2
      Contact( "中间变量".加湿快抽空阀V4输出 )
   END_RUNG wire#w1
   RUNG wire#w2
      Contact( "中间变量".脉动阶段快抽空阀V4输出 )
   END_RUNG wire#w1
   RUNG wire#w2
      Contact( "中间变量".通风阶段快抽空阀V4输出 )
   END_RUNG wire#w1
   RUNG wire#w2
      Contact( "中间变量".紧急脉动快抽阀 )
   END_RUNG wire#w1
   RUNG wire#w2
      Contact( "中间变量".紧急通风快抽空阀 )
   END_RUNG wire#w1
   RUNG wire#w2
      Contact( "中间变量".开门脉动快抽空阀V4 )
   END_RUNG wire#w1
   // the same network as SCL:
   "触摸屏".DO快抽空阀 := ("触摸屏".手动操作1.%X0 AND "触摸屏".手动操作1.%X6) OR (NOT "触摸屏".手动操作1.%X0 AND ("中间变量".预处理快抽空阀V4输出 OR "中间变量".加湿快抽空阀V4输出 OR "中间变量".脉动阶段快抽空阀V4输出 OR "中间变量".通风阶段快抽空阀V4输出 OR "中间变量".紧急脉动快抽阀 OR "中间变量".紧急通风快抽空阀 OR "中间变量".开门脉动快抽空阀V4));
END_REGION

REGION Network 6: 加药阀开V10
   "触摸屏".DO加药阀开 := ("触摸屏".手动操作1.%X0 AND "触摸屏".手动操作1.%X4) OR (NOT "触摸屏".手动操作1.%X0 AND "中间变量".加药阶段V5阀开输出);
   "穿刺初不记录压力值2".TON(IN := "触摸屏".DO加药阀开, PT := T#10S);
END_REGION

REGION Network 7: 加药阀关V10
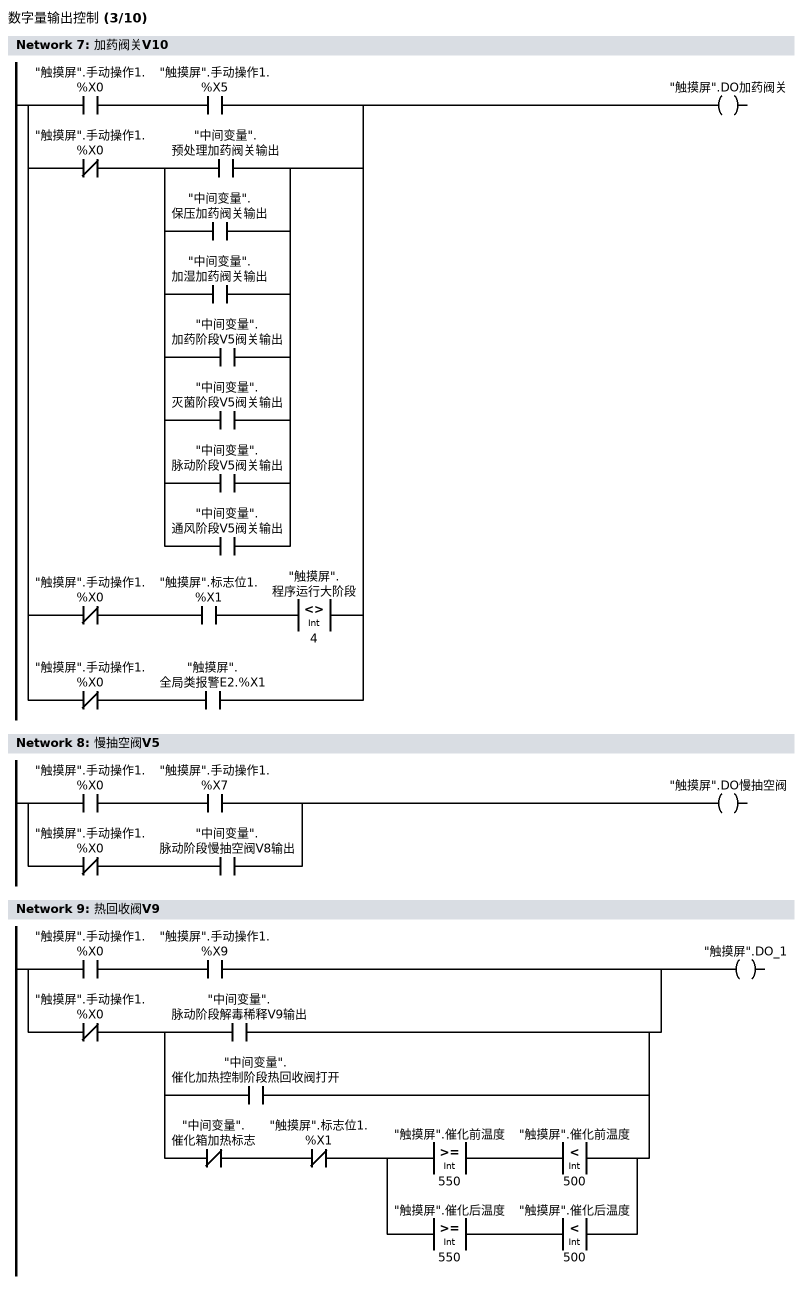
   RUNG wire#powerrail
      Contact( "触摸屏".手动操作1.%X0 )
      Contact( "触摸屏".手动操作1.%X5 )
      wire#w1
      Coil( "触摸屏".DO加药阀关 )
   END_RUNG
   RUNG wire#powerrail
      I_Contact( "触摸屏".手动操作1.%X0 )
      wire#w2
      Contact( "中间变量".预处理加药阀关输出 )
   END_RUNG wire#w1
   RUNG wire#w2
      Contact( "中间变量".保压加药阀关输出 )
   END_RUNG wire#w1
   RUNG wire#w2
      Contact( "中间变量".加湿加药阀关输出 )
   END_RUNG wire#w1
   RUNG wire#w2
      Contact( "中间变量".加药阶段V5阀关输出 )
   END_RUNG wire#w1
   RUNG wire#w2
      Contact( "中间变量".灭菌阶段V5阀关输出 )
   END_RUNG wire#w1
   RUNG wire#w2
      Contact( "中间变量".脉动阶段V5阀关输出 )
   END_RUNG wire#w1
   RUNG wire#w2
      Contact( "中间变量".通风阶段V5阀关输出 )
   END_RUNG wire#w1
   RUNG wire#powerrail
      I_Contact( "触摸屏".手动操作1.%X0 )
      Contact( "触摸屏".标志位1.%X1 )
      { S7_Templates := "SrcType := Int" } NE_Contact(in1 := "触摸屏".程序运行大阶段, in2 := 4)
   END_RUNG wire#w1
   RUNG wire#powerrail
      I_Contact( "触摸屏".手动操作1.%X0 )
      Contact( "触摸屏".全局类报警E2.%X1 )
   END_RUNG wire#w1
   // the same network as SCL:
   "触摸屏".DO加药阀关 := ("触摸屏".手动操作1.%X0 AND "触摸屏".手动操作1.%X5) OR (NOT "触摸屏".手动操作1.%X0 AND ("中间变量".预处理加药阀关输出 OR "中间变量".保压加药阀关输出 OR "中间变量".加湿加药阀关输出 OR "中间变量".加药阶段V5阀关输出 OR "中间变量".灭菌阶段V5阀关输出 OR "中间变量".脉动阶段V5阀关输出 OR "中间变量".通风阶段V5阀关输出)) OR (NOT "触摸屏".手动操作1.%X0 AND "触摸屏".标志位1.%X1 AND ("触摸屏".程序运行大阶段 <> 4)) OR (NOT "触摸屏".手动操作1.%X0 AND "触摸屏".全局类报警E2.%X1);
END_REGION

REGION Network 8: 慢抽空阀V5
   RUNG wire#powerrail
      Contact( "触摸屏".手动操作1.%X0 )
      Contact( "触摸屏".手动操作1.%X7 )
      wire#w1
      Coil( "触摸屏".DO慢抽空阀 )
   END_RUNG
   RUNG wire#powerrail
      I_Contact( "触摸屏".手动操作1.%X0 )
      Contact( "中间变量".脉动阶段慢抽空阀V8输出 )
   END_RUNG wire#w1
   // the same network as SCL:
   "触摸屏".DO慢抽空阀 := ("触摸屏".手动操作1.%X0 AND "触摸屏".手动操作1.%X7) OR (NOT "触摸屏".手动操作1.%X0 AND "中间变量".脉动阶段慢抽空阀V8输出);
END_REGION

REGION Network 9: 热回收阀V9
   RUNG wire#powerrail
      Contact( "触摸屏".手动操作1.%X0 )
      Contact( "触摸屏".手动操作1.%X9 )
      wire#w1
      Coil( "触摸屏".DO_1 )
   END_RUNG
   RUNG wire#powerrail
      I_Contact( "触摸屏".手动操作1.%X0 )
      wire#w2
      Contact( "中间变量".脉动阶段解毒稀释V9输出 )
   END_RUNG wire#w1
   RUNG wire#w2
      Contact( "中间变量".催化加热控制阶段热回收阀打开 )
   END_RUNG wire#w1
   RUNG wire#w2
      I_Contact( "中间变量".催化箱加热标志 )
      I_Contact( "触摸屏".标志位1.%X1 )
      wire#w3
      { S7_Templates := "SrcType := Int" } GE_Contact(in1 := "触摸屏".催化前温度, in2 := 550)
      { S7_Templates := "SrcType := Int" } LT_Contact(in1 := "触摸屏".催化前温度, in2 := 500)
   END_RUNG wire#w1
   RUNG wire#w3
      { S7_Templates := "SrcType := Int" } GE_Contact(in1 := "触摸屏".催化后温度, in2 := 550)
      { S7_Templates := "SrcType := Int" } LT_Contact(in1 := "触摸屏".催化后温度, in2 := 500)
   END_RUNG wire#w1
   // the same network as SCL:
   "触摸屏".DO_1 := ("触摸屏".手动操作1.%X0 AND "触摸屏".手动操作1.%X9) OR (NOT "触摸屏".手动操作1.%X0 AND ("中间变量".脉动阶段解毒稀释V9输出 OR "中间变量".催化加热控制阶段热回收阀打开 OR (NOT "中间变量".催化箱加热标志 AND NOT "触摸屏".标志位1.%X1 AND ((("触摸屏".催化前温度 >= 550) AND ("触摸屏".催化前温度 < 500)) OR (("触摸屏".催化后温度 >= 550) AND ("触摸屏".催化后温度 < 500))))));
END_REGION

REGION Network 10: 催化相关报警，阀的处理
